(* IEC 61131-3 sources: 2026_Projet_YGO_ExcavatriceDragage/CODE/MAIN, 13 files *)

(* ---- GVL_Global.st ---- *)
(* ═══════════════════════════════════════════════════════════════
   🌐 GVL_Global — Variables globales d'utilité générale
   ───────────────────────────────────────────────────────────────
   🎯 Rôle : Regrouper les signaux et horloges système partagés qui
      ne sont pas spécifiques à la logique de simulation ni raccordés
      à des calibrations persistantes.
   ═══════════════════════════════════════════════════════════════ *)
{attribute 'qualified_only'}
VAR_GLOBAL
    BlinkClock1Hz              : BOOL;          // Horloge 1Hz pour clignotements (IHM ou diagnostic)
END_VAR

(* ---- PRG_00_Inputs.st ---- *)
(* ═══════════════════════════════════════════════════════════════
   📥 PRG_00_Inputs — Acquisition et conditionnement des ENTRÉES (PROGRAMME)
   ───────────────────────────────────────────────────────────────
   📄 Doc : DOC/AF_Partie6_IO_Conditioning_v1.2.md §5
   ⚙️ Exécuté par la tâche PLC (Task Manager) en position 0.
   ✅ Expose ses sorties en VAR_OUTPUT (lecture seule pour le reste du code).
   ═══════════════════════════════════════════════════════════════ *)

PROGRAM PRG_00_Inputs
VAR_OUTPUT
    // ── 🛑 SÉCURITÉS COMMUNES (NC — repos=TRUE sain, FALSE=défaut/fil coupé) ──────────────
    // 🔧 REX 2026-07-07 : précision terrain — EmergencyStopOk_DI (retour contact auxiliaire NO)
    // est en fait la confirmation que le CONTACTEUR DE PUISSANCE est réellement engagé (1=actif),
    // PAS la boucle AU elle-même (ça, c'est EmergencyChainOK_DI, ci-dessous). Nom EmergencyStopOk
    // conservé tel quel (contrat FB standard Partie3 §1, utilisé partout) — reste le portail
    // maître du programme, car "puissance réellement présente" est la garantie la plus forte.
    EmergencyStopOk      : BOOL;   // 🚨 Contacteur de puissance confirmé engagé : TRUE=armé/actif ✅ | FALSE=non armé ou coupure 🔴
    EmergencyChain       : BOOL;   // 🔗 REX 2026-07-07 : boucle AU (coup-de-poing + contact PLC) : TRUE=saine ✅ | FALSE=AU appuyé ou PowerCutOff PLC actif 🔴 — précondition à l'armement, PAS le portail maître
    TopPositionSensor    : BOOL;   // 🔝 Fin de course HAUT (NC) : TRUE=libre ✅ | FALSE=butée atteinte 🔴→ForbidAscent
    SlackCableSwitch     : BOOL;   // 🔗 Mou câble sur tambour M2 (NC) : TRUE=câble tendu ✅ | FALSE=mou détecté 🔴→ForbidDescent
    PhaseRotationOk      : BOOL;   // ⚡ Rotation phases élec. (NC) : TRUE=phases OK ✅ | FALSE=inversées/absentes 🔴→SafeStop
    // 🆕 REX 2026-07-08 : retour thermique COMMUN aux 3 freins M1/M2/M3 (1 seul fil, impossible
    // de savoir lequel des 3 est en cause) — demande utilisateur : la perte de ce retour peut
    // signifier un frein qui colle instantanément (frein à manque de courant) → traité comme
    // les autres défauts francs du domaine, escalade PowerCutOff côté FB_Safety_Winch/_Chariot
    // (voir bit10/bit3 respectifs).
    BrakeThermalFeedback : BOOL;   // 🌡️ Thermique frein M1/M2/M3 commun (NC) : TRUE=temp OK ✅ | FALSE=surchauffe ou coupure 🔴→SafeStop+PowerCutOff

    // ── 🪝 TREUIL M1 (frein=NC ; feedback contacteurs=retour unique REX 2026-07-07) ─────
    M1FwdRevSpeedFeedbackOff : BOOL; // 📡 REX 2026-07-07 : retour unique "tous contacteurs (sens+vitesse)
                                      // retombés" M1 — remplace M1ContactorFeedbackFwd/Rev (feedback
                                      // individuel par sens supprimé côté matériel, plus jamais câblé).
                                      // TRUE = tous retombés (sain, rien d'engagé)
    M1ThermalFeedback      : BOOL; // 🌡️ Thermique moteur M1 (NC) : TRUE=temp OK ✅ | FALSE=surchauffe ou coupure 🔴
    M1BrakeFeedback        : BOOL; // 🔒 Retour frein M1 (NC) : TRUE=frein serré repos ✅ | FALSE=desserré/coupure 🔴

    // ── 🪝 TREUIL M2 (même logique que M1) ──────────────────────────────────────────────
    M2FwdRevSpeedFeedbackOff : BOOL; // 📡 REX 2026-07-07 : idem M1, voir ci-dessus
    M2ThermalFeedback      : BOOL; // 🌡️ Thermique moteur M2 (NC) : TRUE=surchauffe ou coupure 🔴→SafeStop+PowerCutOff
    M2BrakeFeedback        : BOOL; // 🔒 Retour frein M2 (NC) : TRUE=serré repos ✅ | FALSE=desserré/coupure 🔴

    // ── ↔️ CHARIOT M3 (capteurs position=NO — position atteinte=TRUE) ────────────────────
    ChariotPosFosse1      : BOOL;  // 📍 Position fosse 1 (NO) : TRUE=chariot en fosse 1 ✅ | FALSE=absent
    ChariotPosFosse2      : BOOL;  // 📍 Position fosse 2 (NO) : TRUE=chariot en fosse 2 ✅ | FALSE=absent
    ChariotPosMaintenance : BOOL;  // 🔧 Position maintenance (NO) : TRUE=en position service ✅ | FALSE=absent
    ChariotPosTremie      : BOOL;  // 🗑️ Position trémie vidange (NO) : TRUE=en position trémie ✅ | FALSE=absent
    M3BrakeFeedback       : BOOL;  // 🔒 Retour frein chariot M3 (NC) : TRUE=serré repos ✅ | FALSE=desserré 🔴

    // 🆕 Variables intermédiaires filtrées/simulées pour contourner la lecture seule des PDO
    M3_StatusWord_Filtered        : WORD;
    M3_ActualFrequencyHz_Filtered : UINT;
END_VAR
VAR
    // Instances de filtrage
    instEmergencyStopOk   : FB_Input;
    instEmergencyChain    : FB_Input; // 🔧 REX 2026-07-07
    instSlackCableSwitch  : FB_Input;
    instTopPositionSensor : FB_Input;
    instCtrlPhaseRotation : FB_Input;
    instBrakeThermalFeedback : FB_Input; // 🆕 REX 2026-07-08

    instM1FwdRevSpeedFeedbackOff : FB_Input; // 🔧 REX 2026-07-07 : remplace instM1ContactorFwd/Rev
    instM1Thermal      : FB_Input;
    instM1BrakeFeedback: FB_Input;

    instM2FwdRevSpeedFeedbackOff : FB_Input; // 🔧 REX 2026-07-07 : remplace instM2ContactorFwd/Rev
    instM2Thermal      : FB_Input;
    instM2BrakeFeedback: FB_Input;

    instChariotPosFosse1      : FB_Input;
    instChariotPosFosse2      : FB_Input;
    instChariotPosMaintenance : FB_Input;
    instChariotPosTremie      : FB_Input;
    instM3BrakeFeedback       : FB_Input;

    // 🧪 Simulation dynamique du trajet chariot M3 (Lot 4, non prioritaire — voir AF_Partie13)
    instSimChariot            : FB_Sim_Chariot;

    // 🧪 Simulation de la chaîne de sécurité AU / réarmement (Lot 1, combler le trou d'intégration)
    instSimSafety             : FB_Sim_Safety;

    // 🧪 Simulation des retours contacteurs et freins M1/M2 (Lot 1)
    M1_FwdRevSpeedFeedbackOff_Simulated : BOOL;
    M1BrakeFeedback_Simulated           : BOOL;
    M2_FwdRevSpeedFeedbackOff_Simulated : BOOL;
    M2BrakeFeedback_Simulated           : BOOL;
    M3BrakeFeedback_Simulated           : BOOL;

    // 🆕 REX 2026-07-08 (4) : cohérence simulation capteur haut (voir instTopPositionSensor ci-dessous)
    SimTopSensorTriggered                : BOOL;
END_VAR

// === IMPLEMENTATION (corps du PROGRAM PRG_00_Inputs) ===

// 🛑 ─── COMMUN ────────────────────────────────────────────────────────────
// 🧪 Simulation : chaque OR ci-dessous force le capteur à son état "sain" (famille
// sécurité, TRUE=OK) quand SimulationModeActive ET que ce capteur précis n'est
// pas encore câblé réellement (GVL_Simulation.*_IsReal). Voir AF_Partie13.

// Simulation de la chaîne de sécurité AU / réarmement (Lot 1)
instSimSafety(
    Enable          := GVL_Simulation.SimulationModeActive AND NOT GVL_Simulation.EmergencyStopChain_IsReal,
    PowerCutOff_A   := PowerCutOff_A_RQ,
    PowerCutOff_B   := PowerCutOff_B_RQ,
    EmergencyArming := EmergencyArming_RQ
);

instEmergencyStopOk(InputRaw := EmergencyStopOk_DI OR instSimSafety.SimContactorOk, FilterTime := T#20MS);
EmergencyStopOk := instEmergencyStopOk.State;

// 🔧 REX 2026-07-07 : boucle AU (coup-de-poing + contact PLC) — distincte du contacteur de
// puissance ci-dessus. Réutilise le même flag simulation (même sous-système physique AU).
instEmergencyChain(InputRaw := EmergencyChainOK_DI OR instSimSafety.SimChainOk, FilterTime := T#20MS);
EmergencyChain := instEmergencyChain.State;

// 🔧 REX 2026-07-07 : M1_M2_SlackCableSwitch_DI → M2_SlackCableSwitch_DI (capteur physiquement
// uniquement sur le tambour M2, le préfixe M1_M2_ ne reflétait pas la réalité du câblage)
instSlackCableSwitch(InputRaw := M2_SlackCableSwitch_DI OR (GVL_Simulation.SimulationModeActive AND NOT GVL_Simulation.SlackCableSwitch_IsReal), FilterTime := T#20MS);
SlackCableSwitch := instSlackCableSwitch.State;

// 🆕 REX 2026-07-08 (4) : cohérence simulation (demande utilisateur) — l'ancien câblage forçait
// TopPositionSensor à TOUJOURS TRUE (sain) en simulation, quelle que soit la position codeur :
// impossible de tester bit5/Méca D (capteur haut) en simulation, il ne se déclenchait JAMAIS.
// Dérivé désormais de la position M1 simulée (référence de l'ensemble, voir FB_Grappin/
// ActiveOffsetM) — 1 cycle de retard (PRG_00 avant PRG_02 dans l'ordre de tâche), négligeable,
// même principe déjà assumé ailleurs (EncoderFaultPresent, GrappinHoldStillActive).
SimTopSensorTriggered := (NOT PRG_04_Modes.instModes.InhibitM1 AND (PRG_02_Encoders.instEncoderScaleM1.CablePosM >= GVL_PERSISTENT.HomingTargetM1_M))
                      OR (NOT PRG_04_Modes.instModes.InhibitM2 AND (PRG_02_Encoders.instEncoderScaleM2.CablePosM >= GVL_PERSISTENT.HomingTargetM2_M));
instTopPositionSensor(InputRaw := M1_M2_TopPositionSensor_DI OR (GVL_Simulation.SimulationModeActive AND NOT GVL_Simulation.TopPositionSensor_IsReal AND NOT SimTopSensorTriggered), FilterTime := T#20MS);
TopPositionSensor := instTopPositionSensor.State;

instCtrlPhaseRotation(InputRaw := CtrlPhaseRotation_DI OR (GVL_Simulation.SimulationModeActive AND NOT GVL_Simulation.PhaseRotationOk_IsReal), FilterTime := T#20MS);
PhaseRotationOk := instCtrlPhaseRotation.State;

// 🆕 REX 2026-07-08 : thermique frein commun M1/M2/M3 (1 seul fil, voir bandeau ci-dessus)
instBrakeThermalFeedback(InputRaw := BrakeThermalFeedback_DI OR (GVL_Simulation.SimulationModeActive AND NOT GVL_Simulation.BrakeThermal_IsReal), FilterTime := T#20MS);
BrakeThermalFeedback := instBrakeThermalFeedback.State;

// 🪝 ─── WINCH M1 ──────────────────────────────────────────────────────────
// 🧪 Simulation des retours contacteurs M1 (retombés si aucun sens/vitesse commandé)
M1_FwdRevSpeedFeedbackOff_Simulated := NOT (PRG_10_Outputs.M1RelayFwd OR PRG_10_Outputs.M1RelayRev OR PRG_10_Outputs.M1SpeedContactor1 OR PRG_10_Outputs.M1SpeedContactor2 OR PRG_10_Outputs.M1SpeedContactor3 OR PRG_10_Outputs.M1SpeedContactor4);
instM1FwdRevSpeedFeedbackOff(InputRaw := SEL(GVL_Simulation.SimulationModeActive AND NOT GVL_Simulation.ContactorFeedbackM1_IsReal, M1_FwdRevSpeedFeedbackOff_DI, M1_FwdRevSpeedFeedbackOff_Simulated), FilterTime := T#20MS);
M1FwdRevSpeedFeedbackOff := instM1FwdRevSpeedFeedbackOff.State;

instM1Thermal(InputRaw := M1_ThermalFeedback_DI OR (GVL_Simulation.SimulationModeActive AND NOT GVL_Simulation.ThermalM1_IsReal), FilterTime := T#20MS);
M1ThermalFeedback := instM1Thermal.State;

// 🧪 Simulation du retour frein M1 (fermé si commande inactive)
M1BrakeFeedback_Simulated := NOT PRG_10_Outputs.M1BrakeCmd;
instM1BrakeFeedback(InputRaw := SEL(GVL_Simulation.SimulationModeActive AND NOT GVL_Simulation.ContactorFeedbackM1_IsReal, M1_BrakeFeedback_DI, M1BrakeFeedback_Simulated), FilterTime := T#20MS);
M1BrakeFeedback := instM1BrakeFeedback.State;

// 🪝 ─── WINCH M2 ──────────────────────────────────────────────────────────
// 🧪 Simulation des retours contacteurs M2 (retombés si aucun sens/vitesse commandé)
M2_FwdRevSpeedFeedbackOff_Simulated := NOT (PRG_10_Outputs.M2RelayFwd OR PRG_10_Outputs.M2RelayRev OR PRG_10_Outputs.M2SpeedContactor1 OR PRG_10_Outputs.M2SpeedContactor2 OR PRG_10_Outputs.M2SpeedContactor3 OR PRG_10_Outputs.M2SpeedContactor4);
instM2FwdRevSpeedFeedbackOff(InputRaw := SEL(GVL_Simulation.SimulationModeActive AND NOT GVL_Simulation.ContactorFeedbackM2_IsReal, M2_FwdRevSpeedFeedbackOff_DI, M2_FwdRevSpeedFeedbackOff_Simulated), FilterTime := T#20MS);
M2FwdRevSpeedFeedbackOff := instM2FwdRevSpeedFeedbackOff.State;

instM2Thermal(InputRaw := M2_ThermalFeedback_DI OR (GVL_Simulation.SimulationModeActive AND NOT GVL_Simulation.ThermalM2_IsReal), FilterTime := T#20MS);
M2ThermalFeedback := instM2Thermal.State;

// 🧪 Simulation du retour frein M2 (fermé si commande inactive)
M2BrakeFeedback_Simulated := NOT PRG_10_Outputs.M2BrakeCmd;
instM2BrakeFeedback(InputRaw := SEL(GVL_Simulation.SimulationModeActive AND NOT GVL_Simulation.ContactorFeedbackM2_IsReal, M2_BrakeFeedback_DI, M2BrakeFeedback_Simulated), FilterTime := T#20MS);
M2BrakeFeedback := instM2BrakeFeedback.State;

// ↔️ ─── CHARIOT M3 ────────────────────────────────────────────────────────
// 🧪 Simulation dynamique du trajet M3 (FB_Sim_Chariot, non prioritaire — voir AF_Partie13
// §Chariot). Appelée AVANT les FB_Input pour que ses sorties soient à jour au même cycle
// (sinon décalage d'1 cycle sur le OR ci-dessous). Remplace le forçage manuel en vue instance.
// 🔧 REX 2026-07-15 (3) : RelayFwd/RelayRev câblés sur M3_CommandWord (variable globale
// mappée PDO EtherCAT, valeur réellement envoyée, Auto ET Manu confondus) — ex-
// GVL_Chariot_M3_Stub.M3_RelayFwd/Rev n'étaient plus jamais écrits depuis l'abandon du mode
// relais DEGRADED_IO (v0.4.11), la simulation de trajet M3 restait bloquée en permanence
// (relais toujours FALSE). Lecture décalée d'1 cycle (10ms, M3_CommandWord réécrit en position
// 10 par PRG_10_Outputs après ce PRG_00) — négligeable devant TravelTimeS (8s).
instSimChariot(
    Enable      := GVL_Simulation.SimulationModeActive AND NOT GVL_Simulation.ChariotPosition_IsReal,
    TargetNum   := GVL_Chariot_M3_Stub.StubChariotPositionSelect_IHM,
    RelayFwd    := M3_CommandWord = 1,
    RelayRev    := M3_CommandWord = 2,
    TravelTimeS := 8.0
);

instChariotPosFosse1(InputRaw := PosFosse1_DI OR instSimChariot.PosFosse1, FilterTime := T#20MS);
ChariotPosFosse1 := instChariotPosFosse1.State;

instChariotPosFosse2(InputRaw := PosFosse2_DI OR instSimChariot.PosFosse2, FilterTime := T#20MS);
ChariotPosFosse2 := instChariotPosFosse2.State;

instChariotPosMaintenance(InputRaw := PosMaintenance_DI OR instSimChariot.PosMaintenance, FilterTime := T#20MS);
ChariotPosMaintenance := instChariotPosMaintenance.State;

instChariotPosTremie(InputRaw := PosTremie_DI OR instSimChariot.PosTremie, FilterTime := T#20MS);
ChariotPosTremie := instChariotPosTremie.State;

// 🧪 Simulation du retour frein M3 (fermé/NC=TRUE si commande inactive)
M3BrakeFeedback_Simulated := NOT PRG_07_ChariotControl.instChariotM3.BrakeCmd;
instM3BrakeFeedback(InputRaw := SEL(GVL_Simulation.SimulationModeActive AND NOT GVL_Simulation.ContactorFeedbackM3_IsReal, M3_BrakeFeedback_DI, M3BrakeFeedback_Simulated), FilterTime := T#20MS);
M3BrakeFeedback := instM3BrakeFeedback.State;

// 🧪 Simulation/Filtrage des retours variateur EtherCAT M3 (lecture seule physique contournée)
IF GVL_Simulation.SimulationModeActive AND NOT GVL_Simulation.VariateurM3_IsReal THEN
    M3_ActualFrequencyHz_Filtered := M3_SetpointFrequencyHz;

    // Status Word : Bit0 (Operation), Bit7 (Operation Enable)
    IF M3_CommandWord = 1 THEN
        M3_StatusWord_Filtered := 16#0081; // Operation + Operation Enable
    ELSIF M3_CommandWord = 2 THEN
        M3_StatusWord_Filtered := 16#0089; // Operation + Operation Enable + Reverse (bit3)
    ELSE
        M3_StatusWord_Filtered := 16#0080; // Stopped + Operation Enable
    END_IF;
ELSE
    M3_ActualFrequencyHz_Filtered := M3_ActualFrequencyHz;
    M3_StatusWord_Filtered        := M3_StatusWord;
END_IF;

(* ---- PRG_01_Diagnostics.st ---- *)
(* ═══════════════════════════════════════════════════════════════
   📡 PRG_01_Diagnostics — États bus de terrain et Joystick (PROGRAMME)
   ───────────────────────────────────────────────────────────────
   ⚙️ Exécuté par la tâche PLC en position 1.
   ═══════════════════════════════════════════════════════════════ *)

PROGRAM PRG_01_Diagnostics
VAR
    instDiagCanOpen  : FB_DiagCanOpen;       // Diagnostic CAN/Joystick
    instDiagEthercat : FB_DiagEthercat;      // Diagnostic EtherCAT (3 devices)
    FB_Joystick_0    : FB_Joystick;          // Traitement joystick (calib/filtre/rampe)
    instSimJoystick  : FB_Sim_Joystick;      // 🧪 Simulation joystick (Lot 3 — voir CODE/SIMULATION/)
END_VAR

// === IMPLEMENTATION (corps du PROGRAM PRG_01_Diagnostics) ===

// 🧪 0. Simulation Joystick (Lot 3, priorité — voir CODE/SIMULATION/FB_Sim_Joystick.st) : appelée
// AVANT FB_Joystick_0 pour que ses sorties soient à jour au même cycle. Remplace l'ancien bypass
// homme-mort codé en dur dans FB_Joystick (GVL_DEBUG.DBG_DeadmanBypass_TEST) : quand
// NOT JoystickSignal_IsReal, ses sorties remplacent les entrées brutes ci-dessous ; le homme-mort
// réel de FB_Joystick n'est plus jamais contourné.
// 🆕 REX 2026-07-08 : gardé désormais par JoystickSignal_IsReal (PAS Joystick_IsReal, qui ne
// couvre que le bus CANopen ci-dessous) — granularité séparée demandée par l'utilisateur : tester
// le signal joystick réel sans dépendre du diagnostic bus/nœud CANopen (encore simulé sain).
instSimJoystick(
    Enable          := GVL_Simulation.SimulationModeActive AND NOT GVL_Simulation.JoystickSignal_IsReal,
    NeutralRaw      := GVL_Simulation.JoystickForceNeutralRaw,
    MaxRaw          := GVL_Simulation.JoystickForceMaxRaw
);

// 1. Diagnostics CANopen — 🆕 REX 2026-07-08 : gardé par Joystick_IsReal UNIQUEMENT (bus/nœud),
// indépendant de JoystickSignal_IsReal (signal brut ci-dessus) — granularité séparée.
instDiagCanOpen(
    Enable := TRUE,
    Reset := PRG_09_Supervision.FaultMachineReset_IHM,
    CanOnline := (CANbus.GetBusState() = 1) OR (GVL_Simulation.SimulationModeActive AND NOT GVL_Simulation.Joystick_IsReal), // 1 = ACTIVE (ou simulation)
    CanOperational := (JOY1_JOYSTICK_MCB560_CO4201A.GetDeviceState() = DEVICE_STATE.RUNNING) OR (GVL_Simulation.SimulationModeActive AND NOT GVL_Simulation.Joystick_IsReal)
);

// 2. Diagnostics EtherCAT (variateur + 2 codeurs)
instDiagEthercat(
    Enable := TRUE,
    Reset := PRG_09_Supervision.FaultMachineReset_IHM,          // 🔑 Bouton général machine
    VariateurWcState := (AC600_ECAT_Drive.GetDeviceState() <> DEVICE_STATE.RUNNING) AND NOT (GVL_Simulation.SimulationModeActive AND NOT GVL_Simulation.VariateurM3_IsReal),
    VariateurSlaveState := SEL((GVL_Simulation.SimulationModeActive AND NOT GVL_Simulation.VariateurM3_IsReal) OR (AC600_ECAT_Drive.GetDeviceState() = DEVICE_STATE.RUNNING), 0, 8),
    EncoderM1WcState := (COD1_CODEUR.GetDeviceState() <> DEVICE_STATE.RUNNING) AND NOT (GVL_Simulation.SimulationModeActive AND NOT GVL_Simulation.EncoderM1_IsReal),
    EncoderM1SlaveState := SEL((GVL_Simulation.SimulationModeActive AND NOT GVL_Simulation.EncoderM1_IsReal) OR (COD1_CODEUR.GetDeviceState() = DEVICE_STATE.RUNNING), 0, 8),
    EncoderM2WcState := (COD2_CODEUR.GetDeviceState() <> DEVICE_STATE.RUNNING) AND NOT (GVL_Simulation.SimulationModeActive AND NOT GVL_Simulation.EncoderM2_IsReal),
    EncoderM2SlaveState := SEL((GVL_Simulation.SimulationModeActive AND NOT GVL_Simulation.EncoderM2_IsReal) OR (COD2_CODEUR.GetDeviceState() = DEVICE_STATE.RUNNING), 0, 8)
);

// 3. Acquisition Joystick — RawX/RawY/RawButton simulés (instSimJoystick) quand NOT JoystickSignal_IsReal
// 🔴🔧 REX 2026-07-07 — TEST BANC UNIQUEMENT, PAS DE VALEUR PRODUCTION :
//    DeadmanRearmTimeout 10s → 5min, NeutralHoldTime 500ms → 1s (confort d'essai, moins de
//    réappuis/traversées à gérer). ⚠️ RÉDUIT RÉELLEMENT LA SÉCURITÉ HOMME-MORT — à repasser
//    impérativement à T#10S / T#500MS (ou retirer ces 2 lignes, le FB reprend ses défauts sûrs)
//    avant toute mise en service réelle avec la machine.
FB_Joystick_0(
    Enable              := TRUE,
    EmergencyStopOk     := PRG_00_Inputs.EmergencyStopOk,
    Reset               := PRG_09_Supervision.FaultMachineReset_IHM,
    Mode                := PRG_04_Modes.instModes.Mode,  // 🆕 REX 2026-07-08 : désarme le homme-mort au changement de mode
    // 🆕 REX 2026-07-08 : PRG_01 (position 1) s'exécute AVANT PRG_06 (position 6) — GrappinBusy lu
    // ici reflète donc le Busy du scan PRÉCÉDENT (retard d'1 scan, ~10ms, sur la détection du front
    // descendant). Sans impact pratique : très inférieur aux temps de réponse frein/contacteurs
    // (100-300ms, voir FB_Brake) — la commande n'a pas le temps de produire un mouvement réel.
    GrappinBusy         := PRG_06_WinchControl.instGrappin.Busy,
    NeutralXMem         := GVL_PERSISTENT.JoystickNeutralX,
    NeutralYMem         := GVL_PERSISTENT.JoystickNeutralY,
    BusCanOpenOP        := instDiagCanOpen.busCanOpen,
    JoystickOP          := instDiagCanOpen.Joystick,
    RawX                := SEL(instSimJoystick.Enable, JoyXRaw_ANA1, instSimJoystick.RawX),
    RawY                := SEL(instSimJoystick.Enable, JoyYRaw_ANA2, instSimJoystick.RawY),
    RawButton           := SEL(instSimJoystick.Enable, JoyBtnRaw, instSimJoystick.RawButton),
    Calibrate           := GVL_IHM.JoystickJOY1.Calibrate,
    InvertX             := FALSE,
    InvertY             := FALSE,
    Deadband            := 10.0,
    FilterTime          := TIME#100ms,
    AccelRate           := 50.0,
    DecelRate           := 150.0,
    // 🛡️ Délais de sécurité Homme-Mort : temporisations courtes (10s/500ms) si joystick réel, longues (5min/1s) si simulé
    DeadmanRearmTimeout := SEL(NOT GVL_Simulation.SimulationModeActive OR GVL_Simulation.JoystickSignal_IsReal, T#5M, T#10S),
    NeutralHoldTime     := SEL(NOT GVL_Simulation.SimulationModeActive OR GVL_Simulation.JoystickSignal_IsReal, T#1S, T#500MS)
);

(* ---- PRG_02_Encoders.st ---- *)
(* ═══════════════════════════════════════════════════════════════
   🧲 PRG_02_Encoders — Acquisition, Recalage (Homing) et Sécurité Codeurs
   ───────────────────────────────────────────────────────────────
   ⚙️ Exécuté par la tâche PLC en position 2.
   ✅ Expose ses défauts en VAR_OUTPUT (1 cycle de retard assumé pour instModes).
   ═══════════════════════════════════════════════════════════════ *)

PROGRAM PRG_02_Encoders
VAR_OUTPUT
    EncoderFaultPresent   : BOOL;   // OR des deux - lu par PRG_04_Modes au cycle suivant
    EncoderFaultPresentM1 : BOOL;
    EncoderFaultPresentM2 : BOOL;
END_VAR
VAR
    // 🧪 Simulation banc de test (Lot 2 — voir CODE/SIMULATION/FB_Sim_Encoder.st)
    instSimEncoderM1      : FB_Sim_Encoder;
    instSimEncoderM2      : FB_Sim_Encoder;
    M1_RawPosToUse        : UDINT;
    M2_RawPosToUse        : UDINT;

    // Instances
    instEncoderAbsM1   : FB_Encoder_Abs;
    instEncoderScaleM1 : FB_Encoder_Scale;
    instHomingM1       : FB_Encoder_Homing;
    instEncoderAbsM2   : FB_Encoder_Abs;
    instEncoderScaleM2 : FB_Encoder_Scale;
    instHomingM2       : FB_Encoder_Homing;
    instEncoderSafetyM1 : FB_Encoder_Safety;
    instEncoderSafetyM2 : FB_Encoder_Safety;

    M1_SimSpeedPct      : REAL;
    M2_SimSpeedPct      : REAL;
    M1_IsReal           : BOOL;         // ⚡ Indique si le treuil M1 est configuré comme réel
    M2_IsReal           : BOOL;         // ⚡ Indique si le treuil M2 est configuré comme réel
END_VAR

// === IMPLEMENTATION (corps du PROGRAM PRG_02_Encoders) ===

// 🆕 Détermination de la réalité des treuils (Conditional Bypass Doctrine)
M1_IsReal := NOT GVL_Simulation.SimulationModeActive OR GVL_Simulation.EncoderM1_IsReal OR GVL_Simulation.ContactorFeedbackM1_IsReal OR GVL_Simulation.ThermalM1_IsReal;
M2_IsReal := NOT GVL_Simulation.SimulationModeActive OR GVL_Simulation.EncoderM2_IsReal OR GVL_Simulation.ContactorFeedbackM2_IsReal OR GVL_Simulation.ThermalM2_IsReal;

// 🔧 REX 2026-07-15 (4) — CORRECTIF COMPILATION : ex-SEL(ManuActive, ...) référençait
// PRG_10_Outputs.SpeedRefPct, supprimé lors du passage de Manu sur FB_Winch (REX 2026-07-15 (2)).
// Plus besoin de distinguer Auto/Manu ici : instWinchM1/M2.SpeedRamp.Current est désormais LA
// vitesse rampée réelle dans les DEUX cas (FB_Winch pilote M1/M2 qu'on soit en Auto ou en Manu).
M1_SimSpeedPct := PRG_06_WinchControl.instWinchM1.SpeedRamp.Current;
M2_SimSpeedPct := PRG_06_WinchControl.instWinchM2.SpeedRamp.Current;

// 1. SIMULATION SUR BANC DE TEST (Lot 2, granularité indépendante M1/M2 — voir AF_Partie13)
// 🔧 REX 2026-07-08 : RawPos (VAR_IN_OUT) référence GVL_PERSISTENT.SimEncoderRawPosM1/M2 —
// survit à un reset froid comme le ferait un vrai codeur absolu physique (voir GVL_PERSISTENT.st).
instSimEncoderM1(
    Enable      := GVL_Simulation.SimulationModeActive AND NOT GVL_Simulation.EncoderM1_IsReal,
    // 🔧 REX 2026-07-15 (2) : lit directement instWinchM1 (PRG_06_WinchControl) — M1 est désormais
    // piloté par FB_Winch en Auto ET en Manu (ex-SimM1Fwd_Eff/PRG_10_Outputs retiré, obsolète) :
    // RelayFwd/RelayRev respectent déjà SafeStop/ForbidAscent/ForbidDescent nativement, plus besoin
    // de signaux Sim dédiés.
    RelayFwd    := PRG_06_WinchControl.instWinchM1.RelayFwd,
    RelayRev    := PRG_06_WinchControl.instWinchM1.RelayRev,
    SpeedRefPct := M1_SimSpeedPct,
    PresetCmd   := (COD1_PresettTrigCmd = 2),
    PresetValue := COD1_PresetValue,
    SpeedScaleFactor := GVL_Simulation.EncoderSimSpeedFactor,  // 🔧 REX 2026-07-07 : confort de test
    // 🆕 REX 2026-07-08 (4) : injection saut de test (Concept 1 / Méca E) — 4096 = PointsPerRev/CableM_PerRev (8192/2.0)
    TestOffsetCmd := GVL_Simulation.InjectSyncDeviationM1,
    TestOffsetPts := REAL_TO_DINT(GVL_Simulation.SyncDeviationOffsetM * 4096.0),
    RawPos      := GVL_PERSISTENT.SimEncoderRawPosM1
);
instSimEncoderM2(
    Enable      := GVL_Simulation.SimulationModeActive AND NOT GVL_Simulation.EncoderM2_IsReal,
    // 🔧 REX 2026-07-15 (2) : idem M1 ci-dessus, lit instWinchM2 (ex-SimM2Fwd_Eff retiré).
    RelayFwd    := PRG_06_WinchControl.instWinchM2.RelayFwd,
    RelayRev    := PRG_06_WinchControl.instWinchM2.RelayRev,
    SpeedRefPct := M2_SimSpeedPct,
    PresetCmd   := (COD2_PresettTrigCmd = 2),
    PresetValue := COD2_PresetValue,
    SpeedScaleFactor := GVL_Simulation.EncoderSimSpeedFactor,  // 🔧 REX 2026-07-07 : confort de test
    // 🆕 REX 2026-07-08 (4) : injection saut de test (Concept 1 / Méca E)
    TestOffsetCmd := GVL_Simulation.InjectSyncDeviationM2,
    TestOffsetPts := REAL_TO_DINT(GVL_Simulation.SyncDeviationOffsetM * 4096.0),
    RawPos      := GVL_PERSISTENT.SimEncoderRawPosM2
);

// Aiguillage (par device — 🔧 REX 2026-07-07 : ne PAS utiliser Operational, forcé à TRUE en
// simulation par PRG_01_Diagnostics [SEL sur EncoderMx_IsReal] pour ne pas remonter de faux
// défaut bus — ça sélectionnait donc systématiquement COD1/COD2_PosValue [réel, figé à 0] au
// lieu de la position simulée, bloquant tout homing/mouvement testé en simulation.
IF (GVL_Simulation.SimulationModeActive AND NOT GVL_Simulation.EncoderM1_IsReal) THEN
    M1_RawPosToUse := instSimEncoderM1.RawPosOut;
ELSE
    M1_RawPosToUse := COD1_PosValue;
END_IF;

IF (GVL_Simulation.SimulationModeActive AND NOT GVL_Simulation.EncoderM2_IsReal) THEN
    M2_RawPosToUse := instSimEncoderM2.RawPosOut;
ELSE
    M2_RawPosToUse := COD2_PosValue;
END_IF;

// 2. TREUIL M1 (Abs → Homing → Scale)
// 🔧 REX 2026-07-07 : Homing appelé AVANT Scale (et non l'inverse) — Scale lit HomingRefRaw en
// entrée ; si Scale s'exécutait avant Homing, un homing réussi au cycle N ne serait répercuté
// sur CablePosM qu'au cycle N+1, alors que instHomingM1.Busy (→ InReferencingMode côté
// FB_Safety_Winch) retombe dès le cycle N — décalage d'1 cycle qui désynchronise le garde-fou
// anti-transition de Méca A (bit7) et provoque un faux déclenchement PowerCutOff au cycle N+1
// (saut de position vu hors fenêtre "référencement en cours"). Homing ne dépend d'aucune sortie
// de Scale (RawPos vient d'instEncoderAbsM1) : aucune dépendance circulaire, réordonnancement sûr.
instEncoderAbsM1(
    Enable              := TRUE,
    Reset               := PRG_09_Supervision.FaultMachineReset_IHM,
    EmergencyStopOk     := PRG_00_Inputs.EmergencyStopOk,
    Mode                := PRG_04_Modes.instModes.Mode,
    RawPosIn            := M1_RawPosToUse,
    AlarmsIn            := SEL(instSimEncoderM1.Enable, COD1_Alarms, 0),
    WarningsIn          := SEL(instSimEncoderM1.Enable, COD1_Warnings, 0),
    SlaveOperational    := PRG_01_Diagnostics.instDiagEthercat.EncoderM1.Operational OR instSimEncoderM1.Enable,
    PresetRequest       := instHomingM1.PresetRequest OR (PRG_10_Outputs.ManuActive AND NOT M1_IsReal AND GVL_IHM.IHM_MANU.HomingEncoder_M1),
    PresetValue         := SEL(PRG_10_Outputs.ManuActive AND NOT M1_IsReal AND GVL_IHM.IHM_MANU.HomingEncoder_M1, instHomingM1.PresetValue, 16777216)
);
COD1_PresettTrigCmd := instEncoderAbsM1.PresetTriggerCmd;
COD1_CodeSeqTrigCmd := instEncoderAbsM1.CodeSeqTriggerCmd;
COD1_PresetValue    := instEncoderAbsM1.PresetValueOut;

instHomingM1(
    Enable               := TRUE,
    Calib                := GVL_PERSISTENT.CalibM1,
    Reset                := PRG_09_Supervision.FaultMachineReset_IHM,
    EmergencyStopOk      := PRG_00_Inputs.EmergencyStopOk,
    Mode                 := PRG_04_Modes.instModes.Mode,
    // ─────────  Début modification IHM_MANU  ─────────
    // 🆕 REX 2026-07-09 : OR avec HomingEncoder_M1 (mise en service urgence) — même FB, mêmes
    // conditions de sécurité (Mode MAINT_N1/N2, arrêt confirmé), aucune nouvelle dérogation.
    Home                 := GVL_IHM.WinchM1.CmdHome OR GVL_IHM.IHM_MANU.HomingEncoder_M1, // 🔧 REX 2026-07-07 : fusion GVL_Encoder_Stub → GVL_IHM
    // ─────────  Fin modification IHM_MANU  ─────────
    ConfirmCoherence     := GVL_IHM.WinchM1.ConfirmCoherence, // 🔧 REX 2026-07-07 : fusion GVL_Encoder_Stub → GVL_IHM
    TopPositionSensor    := PRG_00_Inputs.TopPositionSensor,
    TopSensorPositionM   := GVL_PERSISTENT.HomingTargetM1_M,
    FwdRevSpeedFeedbackOff := PRG_00_Inputs.M1FwdRevSpeedFeedbackOff, // 🔧 REX 2026-07-07
    BrakeFeedback        := PRG_00_Inputs.M1BrakeFeedback,
    RawPos               := instEncoderAbsM1.RawPos,
    EncoderAvailable     := instEncoderAbsM1.EncoderAvailable,
    PresetAck            := instEncoderAbsM1.PresetAck,
    PresetNak            := instEncoderAbsM1.PresetNak,
    PointsPerRev         := 8192,
    MultiTurnRevsMax     := 4096,
    CableM_PerRev        := 2.0
);

instEncoderScaleM1(
    RawPos          := instEncoderAbsM1.RawPos,
    HomingRefRaw    := instHomingM1.HomingRefRaw,
    CableM_PerRev   := 2.0,
    PointsPerRev    := 8192
);

// 3. TREUIL M2 (Abs → Homing → Scale)
instEncoderAbsM2(
    Enable              := TRUE,
    Reset               := PRG_09_Supervision.FaultMachineReset_IHM,
    EmergencyStopOk     := PRG_00_Inputs.EmergencyStopOk,
    Mode                := PRG_04_Modes.instModes.Mode,
    RawPosIn            := M2_RawPosToUse,
    AlarmsIn            := SEL(instSimEncoderM2.Enable, COD2_Alarms, 0),
    WarningsIn          := SEL(instSimEncoderM2.Enable, COD2_Warnings, 0),
    SlaveOperational    := PRG_01_Diagnostics.instDiagEthercat.EncoderM2.Operational OR instSimEncoderM2.Enable,
    PresetRequest       := instHomingM2.PresetRequest OR (PRG_10_Outputs.ManuActive AND NOT M2_IsReal AND GVL_IHM.IHM_MANU.HomingEncoder_M2),
    PresetValue         := SEL(PRG_10_Outputs.ManuActive AND NOT M2_IsReal AND GVL_IHM.IHM_MANU.HomingEncoder_M2, instHomingM2.PresetValue, 16777216)
);
COD2_PresettTrigCmd := instEncoderAbsM2.PresetTriggerCmd;
COD2_CodeSeqTrigCmd := instEncoderAbsM2.CodeSeqTriggerCmd;
COD2_PresetValue    := instEncoderAbsM2.PresetValueOut;

instHomingM2(
    Enable               := TRUE,
    Calib                := GVL_PERSISTENT.CalibM2,
    Reset                := PRG_09_Supervision.FaultMachineReset_IHM,
    EmergencyStopOk      := PRG_00_Inputs.EmergencyStopOk,
    Mode                 := PRG_04_Modes.instModes.Mode,
    // ─────────  Début modification IHM_MANU  ─────────
    // 🆕 REX 2026-07-09 : OR avec HomingEncoder_M2 (mise en service urgence) — même FB, mêmes
    // conditions de sécurité (Mode MAINT_N1/N2, arrêt confirmé), aucune nouvelle dérogation.
    Home                 := GVL_IHM.WinchM2.CmdHome OR GVL_IHM.IHM_MANU.HomingEncoder_M2, // 🔧 REX 2026-07-07 : fusion GVL_Encoder_Stub → GVL_IHM
    // ─────────  Fin modification IHM_MANU  ─────────
    ConfirmCoherence     := GVL_IHM.WinchM2.ConfirmCoherence, // 🔧 REX 2026-07-07 : fusion GVL_Encoder_Stub → GVL_IHM
    TopPositionSensor    := PRG_00_Inputs.TopPositionSensor,
    TopSensorPositionM   := GVL_PERSISTENT.HomingTargetM2_M,
    FwdRevSpeedFeedbackOff := PRG_00_Inputs.M2FwdRevSpeedFeedbackOff, // 🔧 REX 2026-07-07
    BrakeFeedback        := PRG_00_Inputs.M2BrakeFeedback,
    RawPos               := instEncoderAbsM2.RawPos,
    EncoderAvailable     := instEncoderAbsM2.EncoderAvailable,
    PresetAck            := instEncoderAbsM2.PresetAck,
    PresetNak            := instEncoderAbsM2.PresetNak,
    PointsPerRev         := 8192,
    MultiTurnRevsMax     := 4096,
    CableM_PerRev        := 2.0
);

instEncoderScaleM2(
    RawPos          := instEncoderAbsM2.RawPos,
    HomingRefRaw    := instHomingM2.HomingRefRaw,
    CableM_PerRev   := 2.0,
    PointsPerRev    := 8192
);

// 4. SÉCURITÉ DE BORNAGE ET INCOHÉRENCE
instEncoderSafetyM1(
    Enable          := TRUE,
    Reset           := PRG_09_Supervision.FaultMachineReset_IHM,
    EmergencyStopOk := PRG_00_Inputs.EmergencyStopOk,
    Mode            := PRG_04_Modes.instModes.Mode,
    CablePosM       := instEncoderScaleM1.CablePosM,
    HomingSuspect   := instHomingM1.HomingSuspect,
    PositionMinM    := -99.0,
    PositionMaxM    := 99.0
);
EncoderFaultPresentM1 := instEncoderSafetyM1.EncoderIncoherent;

instEncoderSafetyM2(
    Enable          := TRUE,
    Reset           := PRG_09_Supervision.FaultMachineReset_IHM,
    EmergencyStopOk := PRG_00_Inputs.EmergencyStopOk,
    Mode            := PRG_04_Modes.instModes.Mode,
    CablePosM       := instEncoderScaleM2.CablePosM,
    HomingSuspect   := instHomingM2.HomingSuspect,
    PositionMinM    := -99.0,
    PositionMaxM    := 99.0
);
EncoderFaultPresentM2 := instEncoderSafetyM2.EncoderIncoherent;

EncoderFaultPresent := EncoderFaultPresentM1 OR EncoderFaultPresentM2;

// ─────────  Début modification IHM_MANU  ─────────
// 🎯 Référencement direct (bypass sécurité et modes) si HomingEncoder_M1/M2 activés en Manu (uniquement si SIMULÉ)
// Sinon, si les treuils sont réels, on utilise le homing normal sécurisé, et on réinitialise le bouton HMI dès que homing ok/erreur.
IF PRG_10_Outputs.ManuActive THEN
    IF GVL_IHM.IHM_MANU.HomingEncoder_M1 THEN
        IF NOT M1_IsReal THEN
            IF instEncoderAbsM1.PresetAck THEN
                GVL_PERSISTENT.CalibM1.HomingRefRaw := 16726016; // 16777216 - (12.5 * 8192 / 2.0)
                GVL_PERSISTENT.CalibM1.Homed := TRUE;
                GVL_PERSISTENT.CalibM1.HomingSuspect := FALSE;
                GVL_PERSISTENT.CalibM1.LastKnownRawPos := 16777216;
                GVL_IHM.IHM_MANU.HomingEncoder_M1 := FALSE; // Reset bouton HMI
            ELSIF instEncoderAbsM1.PresetNak THEN
                GVL_IHM.IHM_MANU.HomingEncoder_M1 := FALSE;
            END_IF;
        ELSE
            IF instEncoderAbsM1.PresetAck OR instHomingM1.Homed THEN
                GVL_IHM.IHM_MANU.HomingEncoder_M1 := FALSE;
            ELSIF instEncoderAbsM1.PresetNak OR instHomingM1.Error THEN
                GVL_IHM.IHM_MANU.HomingEncoder_M1 := FALSE;
            END_IF;
        END_IF;
    END_IF;

    IF GVL_IHM.IHM_MANU.HomingEncoder_M2 THEN
        IF NOT M2_IsReal THEN
            IF instEncoderAbsM2.PresetAck THEN
                GVL_PERSISTENT.CalibM2.HomingRefRaw := 16726016; // 16777216 - (12.5 * 8192 / 2.0)
                GVL_PERSISTENT.CalibM2.Homed := TRUE;
                GVL_PERSISTENT.CalibM2.HomingSuspect := FALSE;
                GVL_PERSISTENT.CalibM2.LastKnownRawPos := 16777216;
                GVL_IHM.IHM_MANU.HomingEncoder_M2 := FALSE; // Reset bouton HMI
            ELSIF instEncoderAbsM2.PresetNak THEN
                GVL_IHM.IHM_MANU.HomingEncoder_M2 := FALSE;
            END_IF;
        ELSE
            IF instEncoderAbsM2.PresetAck OR instHomingM2.Homed THEN
                GVL_IHM.IHM_MANU.HomingEncoder_M2 := FALSE;
            ELSIF instEncoderAbsM2.PresetNak OR instHomingM2.Error THEN
                GVL_IHM.IHM_MANU.HomingEncoder_M2 := FALSE;
            END_IF;
        END_IF;
    END_IF;
END_IF;
// ─────────  Fin modification IHM_MANU  ─────────

(* ---- PRG_03_Safety.st ---- *)
(* ═══════════════════════════════════════════════════════════════
   🛡️ PRG_03_Safety — Centralisation des surveillances et blocs Safety
   ───────────────────────────────────────────────────────────────
   ⚙️ Exécuté par la tâche PLC en position 3.
   ═══════════════════════════════════════════════════════════════ *)

PROGRAM PRG_03_Safety
VAR
    instSafetyWinchM1   : FB_Safety_Winch;
    instSafetyWinchM2   : FB_Safety_Winch;
    instSafetyChariotM3 : FB_Safety_Chariot;
END_VAR

// === IMPLEMENTATION (corps du PROGRAM PRG_03_Safety) ===

// 1. Sécurité Treuil M1
instSafetyWinchM1(
    // 🔧 REX 2026-07-15 (2) — SIMPLIFICATION : IHM_MANU pilote désormais M1 via FB_Winch
    // (PRG_06_WinchControl), qui a BESOIN d'un SafeStop/ForbidAscent/ForbidDescent réels pour
    // rampé/ralentir proprement (ex-doctrine "Conditional Bypass" devenue obsolète et RETIRÉE
    // ici : chaque capteur/retour a DÉJÀ sa propre granularité réel/simulé — GVL_Simulation.
    // EncoderM1_IsReal, ContactorFeedbackM1_IsReal, ThermalM1_IsReal, TopPositionSensor_IsReal,
    // SlackCableSwitch_IsReal — un composant simulé est déjà forcé "sain" en amont (PRG_00_Inputs/
    // PRG_02_Encoders), donc Enable n'a plus besoin de bypasser tout le domaine : un vrai défaut
    // sur un composant RÉEL protège, un composant SIMULÉ ne fait jamais défaut de lui-même).
    Enable              := NOT PRG_04_Modes.instModes.InhibitM1, // 🆕 REX 2026-07-08 : Inhibit (MAINT_N2) uniquement
    Reset               := PRG_09_Supervision.FaultMachineReset_IHM,
    EmergencyStopOk     := PRG_00_Inputs.EmergencyStopOk,
    Mode                := PRG_04_Modes.instModes.Mode,
    SyncEnable          := PRG_04_Modes.instModes.SyncEnable,
    JoystickOnline      := PRG_01_Diagnostics.instDiagCanOpen.Joystick.Online,
    JoystickOperational := PRG_01_Diagnostics.instDiagCanOpen.Joystick.Operational,
    EncoderAvailable    := PRG_02_Encoders.instEncoderAbsM1.EncoderAvailable,
    ThermalFeedback     := NOT PRG_00_Inputs.M1ThermalFeedback,
    BrakeThermalFeedback := NOT PRG_00_Inputs.BrakeThermalFeedback, // 🆕 REX 2026-07-08 — commun M1/M2/M3
    SlackCableDetected  := NOT PRG_00_Inputs.SlackCableSwitch,
    PhaseRotationOk     := PRG_00_Inputs.PhaseRotationOk,
    TopPositionSensor   := PRG_00_Inputs.TopPositionSensor,
    InReferencingMode   := PRG_02_Encoders.instHomingM1.Busy,
    CablePosM           := PRG_02_Encoders.instEncoderScaleM1.CablePosM,
    CableLimitDescentM  := GVL_PERSISTENT.CableLimitDescentM1_M,
    Direction           := PRG_06_WinchControl.M1_Direction_Active,
    Homed               := PRG_02_Encoders.instHomingM1.Homed,
    HomingSuspect       := PRG_02_Encoders.instHomingM1.HomingSuspect,
    TopLimitM           := GVL_PERSISTENT.HomingTargetM1_M,
    // 🔧 REX 2026-07-07 — Méca A/B/C (voir FB_Safety_Winch bandeau en-tête)
    FwdRevSpeedFeedbackOff := PRG_00_Inputs.M1FwdRevSpeedFeedbackOff,
    BrakeFeedback          := PRG_00_Inputs.M1BrakeFeedback,
    // 🔧 REX 2026-07-15 (7) — BUG CORRIGÉ (retour terrain, SafetyErrorId=256/bit8) : Méca B ne
    // regardait QUE le joystick CANopen pour détecter "commande opérateur" — en IHM_MANU piloté
    // par BOUTONS HMI (JoystickSelect=FALSE), le joystick reste au neutre en permanence, donc
    // MecaB_NoOperatorCmd restait TRUE en continu même pendant un mouvement légitime aux boutons
    // → SafeStop après PostRampTimeout (3s) dès qu'un mouvement HMI dépassait ce délai. Ajout des
    // boutons IHM_MANU bruts (M1 individuel + Couplé) — reste indépendant de l'arbitrage
    // PRG_06/FB_Winch (défense en profondeur intacte, lecture directe des boutons IHM comme le
    // joystick l'était déjà).
    JoystickYNeutral       := (ABS(PRG_01_Diagnostics.FB_Joystick_0.AxisCmdY.SpeedRef) < 0.1)
                              AND NOT GVL_IHM.IHM_MANU.M1_RelayFwd AND NOT GVL_IHM.IHM_MANU.M1_RelayRev
                              AND NOT GVL_IHM.IHM_MANU.M1_M2_RelayFwd AND NOT GVL_IHM.IHM_MANU.M1_M2_RelayRev,
    GrappinHoldStillActive := PRG_06_WinchControl.instGrappin.Busy, // Méca C — M1 doit rester immobile pendant le
                                                                     // grappin ; 1 cycle de retard accepté (PRG_03
                                                                     // avant PRG_06 dans l'ordre de tâche), négligeable
    // 🆕 REX 2026-07-08 (4) — Méca E : M2 corrigé de l'offset grappin actif (0 si grappin absent/ouvert),
    // ramené dans le référentiel M1 — comparaison valable quel que soit l'état du grappin
    ExpectedOtherWinchPosM := PRG_02_Encoders.instEncoderScaleM2.CablePosM - PRG_06_WinchControl.instGrappin.ActiveOffsetM,
    GrappinBusy            := PRG_06_WinchControl.instGrappin.Busy,
    CriticalSyncToleranceM := GVL_PERSISTENT.WinchCriticalSyncTolerance_M,
    OtherWinchInhibited    := PRG_04_Modes.instModes.InhibitM2 // 🆕 REX 2026-07-08 (7)
);

// 2. Sécurité Treuil M2
instSafetyWinchM2(
    // 🔧 REX 2026-07-15 (2) — même simplification que M1 ci-dessus (voir bandeau instSafetyWinchM1).
    Enable              := NOT PRG_04_Modes.instModes.InhibitM2, // 🆕 REX 2026-07-08 : Inhibit (MAINT_N2) uniquement
    Reset               := PRG_09_Supervision.FaultMachineReset_IHM,
    EmergencyStopOk     := PRG_00_Inputs.EmergencyStopOk,
    Mode                := PRG_04_Modes.instModes.Mode,
    SyncEnable          := PRG_04_Modes.instModes.SyncEnable,
    JoystickOnline      := PRG_01_Diagnostics.instDiagCanOpen.Joystick.Online,
    JoystickOperational := PRG_01_Diagnostics.instDiagCanOpen.Joystick.Operational,
    EncoderAvailable    := PRG_02_Encoders.instEncoderAbsM2.EncoderAvailable,
    ThermalFeedback     := NOT PRG_00_Inputs.M2ThermalFeedback,
    BrakeThermalFeedback := NOT PRG_00_Inputs.BrakeThermalFeedback, // 🆕 REX 2026-07-08 — commun M1/M2/M3
    SlackCableDetected  := NOT PRG_00_Inputs.SlackCableSwitch,
    PhaseRotationOk     := PRG_00_Inputs.PhaseRotationOk,
    TopPositionSensor   := PRG_00_Inputs.TopPositionSensor,
    InReferencingMode   := PRG_02_Encoders.instHomingM2.Busy,
    CablePosM           := PRG_02_Encoders.instEncoderScaleM2.CablePosM,
    CableLimitDescentM  := GVL_PERSISTENT.CableLimitDescentM2_M,
    Direction           := PRG_06_WinchControl.M2_Direction_Active,
    Homed               := PRG_02_Encoders.instHomingM2.Homed,
    HomingSuspect       := PRG_02_Encoders.instHomingM2.HomingSuspect,
    TopLimitM           := GVL_PERSISTENT.HomingTargetM2_M,
    // 🔧 REX 2026-07-07 — Méca A/B (voir FB_Safety_Winch bandeau en-tête) — Méca C NON applicable
    // à M2 (c'est M2 qui bouge pendant le grappin, GrappinHoldStillActive reste FALSE)
    FwdRevSpeedFeedbackOff := PRG_00_Inputs.M2FwdRevSpeedFeedbackOff,
    BrakeFeedback          := PRG_00_Inputs.M2BrakeFeedback,
    // 🔧 REX 2026-07-15 (7) : idem M1 (voir bandeau instSafetyWinchM1 ci-dessus).
    JoystickYNeutral       := (ABS(PRG_01_Diagnostics.FB_Joystick_0.AxisCmdY.SpeedRef) < 0.1)
                              AND NOT GVL_IHM.IHM_MANU.M2_RelayFwd AND NOT GVL_IHM.IHM_MANU.M2_RelayRev
                              AND NOT GVL_IHM.IHM_MANU.M1_M2_RelayFwd AND NOT GVL_IHM.IHM_MANU.M1_M2_RelayRev,
    GrappinHoldStillActive := FALSE,
    // 🔧 REX 2026-07-08 (5) : BUG CORRIGÉ — oublié côté M2 lors de l'ajout initial Méca E.
    // ExpectedOtherWinchPosM valait 0.0 par défaut (non câblé) → Méca E comparait CablePosM2
    // à 0 au lieu de M1, déclenchement permanent dès que M2 > CriticalSyncToleranceM (2.0m)
    // du zéro codeur. M1 corrigé de l'offset grappin actif, ramené dans le référentiel M2.
    ExpectedOtherWinchPosM := PRG_02_Encoders.instEncoderScaleM1.CablePosM + PRG_06_WinchControl.instGrappin.ActiveOffsetM,
    GrappinBusy            := PRG_06_WinchControl.instGrappin.Busy,
    CriticalSyncToleranceM := GVL_PERSISTENT.WinchCriticalSyncTolerance_M,
    OtherWinchInhibited    := PRG_04_Modes.instModes.InhibitM1 // 🆕 REX 2026-07-08 (7)
);

// 3. Sécurité Chariot M3
instSafetyChariotM3(
    Enable              := NOT PRG_10_Outputs.ManuActive OR NOT GVL_Simulation.SimulationModeActive OR GVL_Simulation.VariateurM3_IsReal OR GVL_Simulation.ContactorFeedbackM3_IsReal OR GVL_Simulation.ChariotPosition_IsReal, // 🆕 REX 2026-07-14 : ManuActive (Conditional Bypass Doctrine)
    Reset               := PRG_09_Supervision.FaultMachineReset_IHM,
    EmergencyStopOk     := PRG_00_Inputs.EmergencyStopOk,
    Mode                := PRG_04_Modes.instModes.Mode,
    JoystickOnline      := PRG_01_Diagnostics.instDiagCanOpen.Joystick.Online,
    JoystickOperational := PRG_01_Diagnostics.instDiagCanOpen.Joystick.Operational,
    PhaseRotationOk     := PRG_00_Inputs.PhaseRotationOk,
    BrakeThermalFeedback := NOT PRG_00_Inputs.BrakeThermalFeedback, // 🆕 REX 2026-07-08 — commun M1/M2/M3
    DriveOnline         := PRG_01_Diagnostics.instDiagEthercat.Variateur.Online,
    DriveOperational    := PRG_01_Diagnostics.instDiagEthercat.Variateur.Operational,
    DriveStatusWord     := PRG_00_Inputs.M3_StatusWord_Filtered,
    DriveActualFreqHz   := UINT_TO_REAL(PRG_00_Inputs.M3_ActualFrequencyHz_Filtered) / 100.0,
    BrakeFeedback       := PRG_00_Inputs.M3BrakeFeedback,
    BrakeCmd            := PRG_07_ChariotControl.instChariotM3.BrakeCmd,
    Direction           := PRG_07_ChariotControl.M3_Direction_Active,
    LimitSwitchFwd      := PRG_00_Inputs.ChariotPosTremie,
    LimitSwitchRev      := PRG_00_Inputs.ChariotPosFosse1
);

(* ---- PRG_04_Modes.st ---- *)
(* ═══════════════════════════════════════════════════════════════
   🎚️ PRG_04_Modes — Gestion et Arbitrage du Mode Machine
   ───────────────────────────────────────────────────────────────
   ⚙️ Exécuté par la tâche PLC en position 4.
   ═══════════════════════════════════════════════════════════════ *)

PROGRAM PRG_04_Modes
VAR
    instModes : FB_Modes; // Arbitrage du mode machine (DISABLE, MAINT, SEMI_AUTO, etc.)
    PrevInhibitM1 : BOOL; // 🆕 Mémoire d'état M1
    PrevInhibitM2 : BOOL; // 🆕 Mémoire d'état M2
END_VAR

// === IMPLEMENTATION (corps du PROGRAM PRG_04_Modes) ===

// 🆕 Exclusion mutuelle des inhibitions de treuils (soit M1, soit M2, jamais les deux)
IF GVL_IHM.WinchM1.CmdInhibit AND GVL_IHM.WinchM2.CmdInhibit THEN
    // Si M1 était déjà activé, on rejette la demande sur M2 (M2 retombe à FALSE)
    IF PrevInhibitM1 THEN
        GVL_IHM.WinchM2.CmdInhibit := FALSE;
    // Si M2 était déjà activé, on rejette la demande sur M1 (M1 retombe à FALSE)
    ELSIF PrevInhibitM2 THEN
        GVL_IHM.WinchM1.CmdInhibit := FALSE;
    ELSE
        // repli de sécurité si les deux s'activent de façon synchrone sans transition
        GVL_IHM.WinchM1.CmdInhibit := FALSE;
        GVL_IHM.WinchM2.CmdInhibit := FALSE;
    END_IF;
END_IF;

PrevInhibitM1 := GVL_IHM.WinchM1.CmdInhibit;
PrevInhibitM2 := GVL_IHM.WinchM2.CmdInhibit;

// 🆕 Si l'un des treuils est inhibé, synchro impossible par nature -> reset case IHM à TRUE
// (🔧 REX 2026-07-08 : polarité inversée, TRUE = état neutre "synchro voulue")
IF GVL_IHM.WinchM1.CmdInhibit OR GVL_IHM.WinchM2.CmdInhibit THEN
    GVL_IHM.Sync.SyncEnableRequest := TRUE;
END_IF;

instModes(
    Enable              := TRUE,
    Reset               := GVL_IHM.Modes.ModeReset,  // 🔧 REX 2026-07-07 : dédié, jamais mélangé au reset défauts général
    EmergencyStopOk     := PRG_00_Inputs.EmergencyStopOk,
    ModeRequest         := GVL_Modes_Stub.ModeRequest_IHM,      // 🖥️ Sélecteur IHM
    SyncEnableRequest   := GVL_Modes_Stub.SyncEnableRequest_IHM,
    InhibitM1Request    := GVL_IHM.WinchM1.CmdInhibit, // 🆕 REX 2026-07-08 : IHM réelle, pas GVL_Modes_Stub
    InhibitM2Request    := GVL_IHM.WinchM2.CmdInhibit, // 🆕 REX 2026-07-08 : IHM réelle, pas GVL_Modes_Stub
    HomingApproachEnableRequest := GVL_IHM.Common.HomingApproachEnableRequest, // 🆕 REX 2026-07-08 (2)
    EncoderFaultPresent := PRG_02_Encoders.EncoderFaultPresent,   // 1 cycle de retard (reçu de PRG_02_Encoders)
    JoystickWinchSelectRequest := GVL_IHM.IHM_MANU.JoystickWinchSelect // 🆕 TASK-0001
);

(* ---- PRG_05_Cycle.st ---- *)
(* ═══════════════════════════════════════════════════════════════
   🔄 PRG_05_Cycle — Séquenceur du Cycle Automatique / Semi-Auto (Grafcet)
   ───────────────────────────────────────────────────────────────
   ⚙️ Exécuté par la tâche PLC en position 5.
   ✅ Gère la machine d'état principale de dragage (FB_Cycle).
   ═══════════════════════════════════════════════════════════════ *)

PROGRAM PRG_05_Cycle
VAR
    // Instance du séquenceur automatique
    instCycle           : FB_Cycle;

    // Commandes issues de la supervision (IHM)
    CmdStartCycle_IHM   : BOOL;         // Lancement cycle automatique
    CmdPauseCycle_IHM   : BOOL;         // Pause cycle automatique
    CmdAbortCycle_IHM   : BOOL;         // Abandon / arrêt cycle automatique
    CmdResetCycle_IHM   : BOOL;         // 🔧 REX 2026-07-07 : reset dédié FB_Cycle, jamais mélangé au reset défauts général

    // Paramètres cibles réglés par l'opérateur
    TargetDepthM        : REAL := -12.5; // Profondeur de dragage cible (mètres, négative)
    TargetOffsetM       : REAL := 1.5;  // Décalage cible de fermeture du grappin (mètres)
END_VAR

// === IMPLEMENTATION (corps du PROGRAM PRG_05_Cycle) ===

// Appel du séquenceur de cycle principal avec tous ses raccordements
instCycle(
    Enable              := (PRG_04_Modes.instModes.Mode = E_Mode.SEMI_AUTO) AND NOT PRG_10_Outputs.ManuActive,
    Reset               := CmdResetCycle_IHM,
    EmergencyStopOk     := PRG_00_Inputs.EmergencyStopOk,

    StartCycle          := CmdStartCycle_IHM,
    PauseCycle          := CmdPauseCycle_IHM,
    AbortCycle          := CmdAbortCycle_IHM,

    TargetDepthM        := TargetDepthM,
    TargetOffsetM       := TargetOffsetM,
    SelectedTargetNum_IHM := GVL_IHM.ChariotM3.SelectedTargetNum,

    // Capteur fond touché détecté par le mou de câble physique (sécurité positive)
    BottomTouched       := NOT PRG_00_Inputs.SlackCableSwitch,
    M1_CablePosM        := PRG_02_Encoders.instEncoderScaleM1.CablePosM,
    M2_CablePosM        := PRG_02_Encoders.instEncoderScaleM2.CablePosM,

    // Position chariot
    Chariot_At_Fosse1   := PRG_00_Inputs.ChariotPosFosse1,
    Chariot_At_Fosse2   := PRG_00_Inputs.ChariotPosFosse2,
    Chariot_At_Maintenance := PRG_00_Inputs.ChariotPosMaintenance,
    Chariot_At_Tremie   := PRG_00_Inputs.ChariotPosTremie,
    Chariot_Busy        := PRG_07_ChariotControl.instChariotM3.Busy,
    Chariot_Done        := PRG_07_ChariotControl.instChariotM3.Done,

    // Mouvements mâchoires grappin (gérés par instGrappin)
    Grappin_Busy        := PRG_06_WinchControl.instGrappin.Busy,
    Grappin_Done        := PRG_06_WinchControl.instGrappin.Done,
    Grappin_IsOpen      := GVL_PERSISTENT.GrappinState.IsOpen,
    Grappin_IsClosed    := GVL_PERSISTENT.GrappinState.IsClosed
);

(* ---- PRG_06_WinchControl.st ---- *)
(* ═══════════════════════════════════════════════════════════════
   🪝 PRG_06_WinchControl — Commande des Treuils M1/M2, Synchro et Grappin
   ───────────────────────────────────────────────────────────────
   ⚙️ Exécuté par la tâche PLC en position 6.
   ✅ Arbitre entre les commandes Manuelles (Joystick) et Automatiques (PRG_05_Cycle).
   ═══════════════════════════════════════════════════════════════ *)

PROGRAM PRG_06_WinchControl
VAR
    // Stubs
    StubMachineEnableN1 : BOOL := TRUE;

    // Instances
    instWinchSync : FB_WinchSync;
    instGrappin   : FB_Grappin;
    instWinchM1   : FB_Winch;
    instWinchM2   : FB_Winch;

    // Variables de commande M1 après arbitrage Manuel/Auto
    M1_StartStop_Active     : BOOL;
    M1_Direction_Active     : INT;
    M1_SpeedRef_Active      : REAL;

    // Variables de commande M2 après arbitrage Grappin/Manuel/Auto
    M2_StartStop_Active     : BOOL;
    M2_Direction_Active     : INT;
    M2_SpeedRef_Active      : REAL;
    M2_SpeedStepTableActive : ST_SpeedStepTable;

    // Bornage et limites
    BottomLimitM1_Active    : REAL;
    BottomLimitM2_Active    : REAL;
    ForbidDescentM1_Active  : BOOL;
    ForbidDescentM2_Active  : BOOL;
    // 🆕 REX 2026-07-15 (8) — miroir IHM dédié CableLimitAscentM1/2_M (demande utilisateur, symétrique
    // à CableLimitDescentReached) : indique PRÉCISÉMENT que la nouvelle limite haute d'exploitation
    // normale est atteinte (hors capteur physique bit5, hors Homing) — voir §5 plus bas.
    CableLimitAscentM1Reached : BOOL;
    CableLimitAscentM2Reached : BOOL;

    // 🔧 REX 2026-07-07 : couplage croisé M1/M2 des arrêts, UNIQUEMENT si SyncActive (mouvement
    // coherent voulu). Hors synchro (Grappin.Busy ou SyncEnable=FALSE MAINT_N2) : chaque treuil réagit
    // à SA PROPRE limite/défaut uniquement — commande indépendante voulue dans ce cas.
    SafeStopM1_Raw          : BOOL;
    SafeStopM2_Raw          : BOOL;
    SafeStopM1_Active       : BOOL;
    SafeStopM2_Active       : BOOL;
    ForbidDescentM1_Raw     : BOOL;
    ForbidDescentM2_Raw     : BOOL;
    ForbidAscentM1_Raw      : BOOL;
    ForbidAscentM2_Raw      : BOOL;
    ForbidAscentM1_Active   : BOOL;
    ForbidAscentM2_Active   : BOOL;

    // 🆕 REX 2026-07-08 : voir §2bis — coupure immédiate M1/M2 au même scan que la fin du cycle
    // grappin (contrairement au désarmement homme-mort côté FB_Joystick, qui a 1 scan de retard
    // structurel — PRG_01 s'exécute avant PRG_06). Corrige un bref "blip" de commande (RelayFwd/Rev
    // + BrakeCmd clignotant) observé sur M1 à l'arrivée en position grappin.
    GrappinBusyFallEdge     : F_TRIG;

    // 🆕 REX 2026-07-08 (4) : instWinchSync appelé APRÈS l'arbitrage M1/M2 (§3, plus bas) — lu ici
    // avec 1 scan de retard (~10ms), négligeable vu que DeltaPosM évolue progressivement, pas
    // par à-coup (même raisonnement que M1_Busy/M2_Busy sur instGrappin, voir §0).
    SyncMinorDeviation      : BOOL;
    SyncMinorDeviationBlocksUp   : BOOL;   // 🆕 REX 2026-07-08 (5) : bit0 latché ET écart actuel aggravé par la montée
    SyncMinorDeviationBlocksDown : BOOL;   // 🆕 REX 2026-07-08 (5) : bit0 latché ET écart actuel aggravé par la descente
    M2_LimitShift                : REAL;   // 🆕 REX 2026-07-08 : décalage dynamique de la butée haute de M2

    // 🆕 REX 2026-07-15 (3) — demande utilisateur : les fins de course virtuelles grappin
    // (FdcGrappinOpen/CloseActive) doivent bloquer le mouvement AUSSI en pilotage COUPLÉ IHM_MANU
    // (M1+M2 simultané), pas seulement en pilotage individuel M2 — sinon un opérateur qui pousse le
    // couplage alors que le grappin est déjà en butée virtuelle n'est protégé que par la butée
    // mécanique passive. Masque calculé UNE FOIS ici, consommé par M1 ET M2 (§1/§2 ci-dessous) pour
    // que les deux treuils s'arrêtent ENSEMBLE (pas de désynchro M1/M2 en cas de blocage partiel).
    CoupledFwdGrappinOk          : BOOL;   // Couplage montée autorisé (pas de butée fermeture grappin)
    CoupledRevGrappinOk          : BOOL;   // Couplage descente autorisé (pas de butée ouverture grappin)

    // 🆕 REX 2026-07-15 (9) — plafond palier IHM_MANU "essais progressifs" (demande utilisateur,
    // TEMPORAIRE tant que les vitesses définitives ne sont pas figées, à retirer ensuite) : commun
    // aux 2 treuils (GVL_IHM.IHM_MANU.WinchMaxStepFwd/Rev, structure figée, un seul réglage pour M1
    // ET M2). Actif UNIQUEMENT si ManuActive — Auto garde son comportement inchangé (5 en montée,
    // WinchMaxStepDescente en descente). En Manu, le plafond descente est le MIN avec
    // WinchMaxStepDescente (jamais moins protecteur qu'Auto, juste potentiellement plus prudent).
    ManuMaxStepFwd            : INT;
    ManuMaxStepRev            : INT;
    EffectiveMaxStepAscent    : INT;
    EffectiveMaxStepDescente  : INT;
END_VAR

// === IMPLEMENTATION (corps du PROGRAM PRG_06_WinchControl) ===

// ── 0. COMMANDE DU GRAPPIN (Séquence lente) ─────────────────────────────
// 🔧 REX 2026-07-08 : appelé EN PREMIER (avant l'arbitrage M1/M2 ci-dessous) — audit sécurité :
// l'ancien ordre (Grappin appelé après l'arbitrage) faisait que M1_StartStop_Active lisait
// instGrappin.Busy du scan PRÉCÉDENT, créant une fenêtre d'1 scan où M1 pouvait recevoir une
// commande manuelle au moment exact où le grappin démarre. instGrappin.M1_Busy/M2_Busy (ci-dessous)
// lisent en retour instWinchM1/M2.Busy du scan précédent (ces FB sont appelés plus loin, §6/§7) —
// acceptable : ça ne retarde que l'ACCEPTATION d'une nouvelle demande de ~1 scan (10ms), sans
// aucun impact sécurité (contrairement au cas inverse, qui pouvait faire bouger M1 pendant Busy).
instGrappin(
    Enable              := NOT PRG_04_Modes.instModes.InhibitM2
                           AND PRG_02_Encoders.instEncoderAbsM1.EncoderAvailable
                           AND PRG_02_Encoders.instEncoderAbsM2.EncoderAvailable, // 🆕 Sécurisé : nécessite les deux codeurs valides et M2 non-inhibé
    Reset               := PRG_09_Supervision.FaultMachineReset_IHM,
    EmergencyStopOk     := PRG_00_Inputs.EmergencyStopOk,
    Mode                := PRG_04_Modes.instModes.Mode,
    CmdOpen_IHM         := GVL_IHM.Grappin.CmdOpen OR PRG_05_Cycle.instCycle.CmdGrappin_Open,
    CmdClose_IHM        := GVL_IHM.Grappin.CmdClose OR PRG_05_Cycle.instCycle.CmdGrappin_Close,
    JoystickY_StartStop := PRG_01_Diagnostics.FB_Joystick_0.AxisCmdY.StartStop,
    JoystickY_Direction := PRG_01_Diagnostics.FB_Joystick_0.AxisCmdY.Direction,
    CablePosM1          := PRG_02_Encoders.instEncoderScaleM1.CablePosM,
    CablePosM2          := PRG_02_Encoders.instEncoderScaleM2.CablePosM,
    HomedM1             := PRG_02_Encoders.instHomingM1.Homed,
    HomedM2             := PRG_02_Encoders.instHomingM2.Homed,
    M1_Busy             := instWinchM1.Busy,   // 🆕 REX 2026-07-08
    M2_Busy             := instWinchM2.Busy,   // 🆕 REX 2026-07-08
    ConfirmOpenPosition := GVL_IHM.Grappin.CmdConfirmOpenPosition, // 🆕 REX 2026-07-08 — bouton IHM référencement grappin ouvert
    ConfirmClosePosition:= GVL_IHM.Grappin.CmdConfirmClosePosition, // 🆕 REX 2026-07-08 — bouton IHM référencement grappin fermé
    Config              := GVL_PERSISTENT.GrappinConfig,
    TimeoutDuration     := GVL_IHM.Grappin.TimeoutDuration,
    GrappinState        := GVL_PERSISTENT.GrappinState,
    InhibitM1           := PRG_04_Modes.instModes.InhibitM1, // 🆕 REX 2026-07-08
    InhibitM2           := PRG_04_Modes.instModes.InhibitM2  // 🆕 REX 2026-07-08
);

// 🆕 REX 2026-07-08 (4) — Concept 1 (écart synchro mineur) : bit0 seul (écart position, hors
// incohérence commande bit1) ne fait plus de SafeStop (fast) — bloque StartStop → rampe de décél
// NORMALE. Recalage : voir SyncEnable=FALSE (MAINT_N2), procédure déjà existante (mou de câble).
SyncMinorDeviation := (instWinchSync.ErrorId AND 16#0001) <> 16#0000;

// 🔧 REX 2026-07-08 (5) — audit sécurité : ne bloque plus StartStop dans les 2 sens (déblocage
// impossible sans Reset+MAINT_N2, régression terrain constatée, écart mécanique transitoire
// normal à l'arrêt). SignedDeltaPosM > 0 = M1 plus "haut" que M2 : la montée (Direction=+1)
// aggrave cet écart, la descente (-1) le réduit — et inversement si < 0. Seul le sens aggravant
// reste bloqué ; Méca E (FB_Safety_Winch, écart critique 2.0m) et bit1 (incohérence commande)
// restent le filet réel si l'écart continue de dériver malgré cette autorisation directionnelle.
// 🆕 REX 2026-07-08 (6) : gate global SyncSoftStopEnable — FALSE (défaut) = ces 2 sorties
// restent FALSE en permanence (bit0 déjà géré en SafeStop fast classique ci-dessus, §5bis) ;
// TRUE = active le blocage directionnel (nouvelle fonctionnalité, opt-in).
SyncMinorDeviationBlocksUp   := GVL_PERSISTENT.SyncSoftStopEnable AND SyncMinorDeviation AND (instWinchSync.SignedDeltaPosM > 0.0);
SyncMinorDeviationBlocksDown := GVL_PERSISTENT.SyncSoftStopEnable AND SyncMinorDeviation AND (instWinchSync.SignedDeltaPosM < 0.0);

// 🆕 REX 2026-07-15 (3) — voir déclaration VAR ci-dessus : couplé masqué par les mêmes fins de
// course grappin que l'individuel M2, appliqué à M1 ET M2 (§1/§2) pour arrêter les DEUX treuils
// ensemble plutôt que de désynchroniser M1/M2 en ne bloquant que la moitié du couplage.
CoupledFwdGrappinOk := NOT GVL_IHM.IHM_MANU.FdcGrappinCloseActive;
CoupledRevGrappinOk := NOT GVL_IHM.IHM_MANU.FdcGrappinOpenActive;

// 🆕 REX 2026-07-15 (9) — plafond palier IHM_MANU "essais progressifs" (voir déclaration VAR
// ci-dessus). Bornage identique à l'ex-logique PRG_10_Outputs retirée lors du passage sur FB_Winch.
ManuMaxStepFwd := GVL_IHM.IHM_MANU.WinchMaxStepFwd;
IF (ManuMaxStepFwd < 1) OR (ManuMaxStepFwd > 5) THEN
    ManuMaxStepFwd := 5; // Pleine vitesse par défaut si non initialisé/invalide
END_IF;
ManuMaxStepRev := GVL_IHM.IHM_MANU.WinchMaxStepRev;
IF (ManuMaxStepRev < 1) OR (ManuMaxStepRev > 5) THEN
    ManuMaxStepRev := 2; // Palier 2 max par défaut en descente (conforme AF) si non initialisé/invalide
END_IF;
EffectiveMaxStepAscent   := SEL(PRG_10_Outputs.ManuActive, 5, ManuMaxStepFwd);
EffectiveMaxStepDescente := SEL(PRG_10_Outputs.ManuActive, GVL_PERSISTENT.WinchMaxStepDescente, MIN(GVL_PERSISTENT.WinchMaxStepDescente, ManuMaxStepRev));

// ── 1. ARBITRAGE DES CONSIGNES M1 (Joystick vs Cycle Automatique) ────────
IF PRG_04_Modes.instModes.Mode = E_Mode.SEMI_AUTO THEN
    // 🔧 REX 2026-07-08 (7) — review : gate directionnel absent de cette branche (bug trouvé en
    // review code), le cycle auto pouvait aggraver un écart mineur sans aucune protection quand
    // SyncSoftStopEnable=TRUE. Ajouté ici, symétrique à la branche manuelle ci-dessous.
    M1_Direction_Active := PRG_05_Cycle.instCycle.CmdWinchM1_Direction;
    M1_StartStop_Active := PRG_05_Cycle.instCycle.CmdWinchM1_StartStop
                            AND NOT ((SyncMinorDeviationBlocksUp   AND (M1_Direction_Active = 1))
                                 OR  (SyncMinorDeviationBlocksDown AND (M1_Direction_Active = -1)));
    M1_SpeedRef_Active  := PRG_05_Cycle.instCycle.CmdWinchM1_SpeedPct;
ELSIF PRG_10_Outputs.ManuActive THEN
    // 🆕 REX 2026-07-15 (2) — IHM_MANU pilote désormais M1 via FB_Winch (au lieu de l'ex-bypass
    // direct dans PRG_10_Outputs) : récupère gratuitement la rampe accel/décel + le ralentissement
    // en zone d'approche de bordure + le maintien du relais pendant la décél (mêmes paramètres
    // persistants qu'en Auto, voir instWinchM1 plus bas §6). Demande (boutons IHM ou joystick, déjà
    // arbitrée par PRG_10_Outputs : M1Fwd_Demand/M1Rev_Demand/CoupledFwd_Demand/CoupledRev_Demand)
    // lue avec 1 scan de retard (~10ms, PRG_10 position 10 > PRG_06 position 6) — même principe
    // déjà accepté ailleurs dans ce fichier (Grappin.Busy, SyncMinorDeviation).
    // 🔧 REX 2026-07-15 (5) — trouvé en revue croisée (agent Haiku + relecture manuelle) : M1
    // INDIVIDUEL (bouton M1_RelayFwd/Rev, indépendant de M2) n'était masqué par AUCUNE butée
    // grappin — delta = CablePosM1 - CablePosM2, donc bouger M1 seul aggrave la MÊME sur-contrainte
    // mécanique que le couplé (déjà corrigé ci-dessous) : M1 Fwd augmente le delta (aggrave
    // FdcGrappinOpenActive, delta déjà >= 0) ; M1 Rev diminue le delta (aggrave
    // FdcGrappinCloseActive, delta déjà <= -10). Sens INVERSÉ par rapport à M2 (M2Fwd↔Close,
    // M2Rev↔Open) car M1 et M2 ont un effet opposé sur le même delta. Couplé masqué par
    // CoupledFwdGrappinOk/CoupledRevGrappinOk (REX 2026-07-15 (3)) — M1 s'arrête EN MÊME TEMPS que
    // M2 si le couplage OU son propre individuel violerait une butée grappin.
    IF (PRG_10_Outputs.M1Fwd_Demand AND NOT GVL_IHM.IHM_MANU.FdcGrappinOpenActive) OR (PRG_10_Outputs.CoupledFwd_Demand AND CoupledFwdGrappinOk) THEN
        M1_Direction_Active := 1;
    ELSIF (PRG_10_Outputs.M1Rev_Demand AND NOT GVL_IHM.IHM_MANU.FdcGrappinCloseActive) OR (PRG_10_Outputs.CoupledRev_Demand AND CoupledRevGrappinOk) THEN
        M1_Direction_Active := -1;
    ELSE
        M1_Direction_Active := 0;
    END_IF;
    M1_StartStop_Active := (M1_Direction_Active <> 0);
    // 🎯 Joystick = vitesse proportionnelle à la déflexion (comme en Auto) ; boutons HMI = cible 100%
    // (FB_Winch rampe déjà en interne, plus besoin de la rampe HMI locale ex-PRG_10_Outputs).
    M1_SpeedRef_Active  := SEL(GVL_IHM.IHM_MANU.JoystickSelect, 100.0, ABS(PRG_01_Diagnostics.FB_Joystick_0.AxisCmdY.SpeedRef));
ELSE
    // 🔧 REX 2026-07-08 : + AND DeadmanArmed — NOT Busy seul insuffisant (rampe joystick met du
    // temps à redescendre à 0 après désarmement homme-mort ⇒ StartStop reste TRUE le temps de la
    // décél, M1 bougeait/frein décollait à la fin d'un cycle grappin). DeadmanArmed reste FALSE
    // en continu jusqu'au repassage neutre + réappui, sans dépendre du temps de rampe.
    // 🔧 REX 2026-07-08 (5) : Direction assignée AVANT StartStop (nécessaire pour le gate directionnel ci-dessous).
    M1_Direction_Active := PRG_01_Diagnostics.FB_Joystick_0.AxisCmdY.Direction;
    M1_StartStop_Active := PRG_01_Diagnostics.FB_Joystick_0.AxisCmdY.StartStop AND NOT instGrappin.Busy
                            AND PRG_01_Diagnostics.FB_Joystick_0.DeadmanArmed
                            AND NOT ((SyncMinorDeviationBlocksUp   AND (M1_Direction_Active = 1))
                                 OR  (SyncMinorDeviationBlocksDown AND (M1_Direction_Active = -1))); // 🔧 REX 2026-07-08 (5)
    M1_SpeedRef_Active  := PRG_01_Diagnostics.FB_Joystick_0.AxisCmdY.SpeedRef;
END_IF;

// ── 2. ARBITRAGE DES CONSIGNES M2 (Grappin vs Cycle Automatique vs Joystick) ──
IF instGrappin.Busy THEN
    M2_StartStop_Active := instGrappin.M2_StartStop;
    M2_Direction_Active := instGrappin.M2_Direction;
    M2_SpeedRef_Active  := 15.0; // Vitesse lente forcée pour fermeture grappin
ELSE
    IF PRG_04_Modes.instModes.Mode = E_Mode.SEMI_AUTO THEN
        // 🔧 REX 2026-07-08 (7) — review : gate directionnel absent de cette branche, ajouté
        // symétrique à la branche manuelle ci-dessous (signe M2, voir note ci-dessous).
        M2_Direction_Active := PRG_05_Cycle.instCycle.CmdWinchM2_Direction;
        M2_StartStop_Active := PRG_05_Cycle.instCycle.CmdWinchM2_StartStop
                                AND NOT ((SyncMinorDeviationBlocksUp   AND (M2_Direction_Active = -1))
                                     OR  (SyncMinorDeviationBlocksDown AND (M2_Direction_Active = 1)));
        M2_SpeedRef_Active  := PRG_05_Cycle.instCycle.CmdWinchM2_SpeedPct;
    ELSIF PRG_10_Outputs.ManuActive THEN
        // 🔧 REX 2026-07-15 (3) — idem M1 (voir §1) : Fins de course grappin (FdcGrappin) appliquées
        // au pilotage INDIVIDUEL **ET** COUPLÉ de M2 désormais (demande utilisateur — "que ce soit
        // couplé ou pas couplé, il faut rester dans les butées"). Ex-comportement (couplé non
        // masqué) retiré : c'était une incohérence, pas un choix voulu.
        IF (PRG_10_Outputs.M2Fwd_Demand AND NOT GVL_IHM.IHM_MANU.FdcGrappinCloseActive) OR (PRG_10_Outputs.CoupledFwd_Demand AND CoupledFwdGrappinOk) THEN
            M2_Direction_Active := 1;
        ELSIF (PRG_10_Outputs.M2Rev_Demand AND NOT GVL_IHM.IHM_MANU.FdcGrappinOpenActive) OR (PRG_10_Outputs.CoupledRev_Demand AND CoupledRevGrappinOk) THEN
            M2_Direction_Active := -1;
        ELSE
            M2_Direction_Active := 0;
        END_IF;
        M2_StartStop_Active := (M2_Direction_Active <> 0);
        M2_SpeedRef_Active  := SEL(GVL_IHM.IHM_MANU.JoystickSelect, 100.0, ABS(PRG_01_Diagnostics.FB_Joystick_0.AxisCmdY.SpeedRef));
    ELSE
        // 🔧 REX 2026-07-08 : + AND DeadmanArmed, même raison que M1 ci-dessus
        // 🔧 REX 2026-07-08 (5) : Direction assignée AVANT StartStop (gate directionnel)
        // 🐛 REX 2026-07-08 (7) — BUG CORRIGÉ (review code) : signe inversé pour M2. SignedDeltaPosM
        // (référentiel M1 : CablePosM1-CablePosM2+Offset) > 0 signifie M1 en avance — pour RATTRAPER,
        // M2 doit MONTER (+1), pas descendre. Donc BlocksUp (écart M1-en-avance) doit bloquer côté M2
        // le sens qui AGGRAVE, c-à-d Direction=-1 (descendre, M2 prend encore plus de retard) — PAS
        // Direction=+1 (monter, qui RATTRAPE). Symétrique inversé par rapport à M1 (qui utilise +1/-1
        // directement car SignedDeltaPosM est déjà dans SON référentiel).
        M2_Direction_Active := PRG_01_Diagnostics.FB_Joystick_0.AxisCmdY.Direction;
        M2_StartStop_Active := PRG_01_Diagnostics.FB_Joystick_0.AxisCmdY.StartStop
                                AND PRG_01_Diagnostics.FB_Joystick_0.DeadmanArmed
                                AND NOT ((SyncMinorDeviationBlocksUp   AND (M2_Direction_Active = -1))
                                     OR  (SyncMinorDeviationBlocksDown AND (M2_Direction_Active = 1))); // 🔧 REX 2026-07-08 (7)
        M2_SpeedRef_Active  := PRG_01_Diagnostics.FB_Joystick_0.AxisCmdY.SpeedRef;
    END_IF;
END_IF;

// ── 2bis. COUPURE IMMÉDIATE M1/M2 AU SCAN EXACT DE FIN DE CYCLE GRAPPIN ─────
// 🆕 REX 2026-07-08 : instGrappin est appelé en premier (§0), donc son Busy est frais dans CE scan
// (voir §1/§2 ci-dessus) — mais AxisCmdY.StartStop/Direction viennent de FB_Joystick_0 (PRG_01),
// calculé AVANT ce scan de PRG_06. Le désarmement homme-mort sur front descendant de Grappin.Busy
// (FB_Joystick §4ter-ter) ne prend donc effet qu'au scan SUIVANT (~10ms de retard structurel). Si
// l'opérateur tient encore le manche poussé au moment exact où le grappin termine, M1 ET M2
// recevaient pendant ce scan la commande manche brute (RelayFwd/Rev + BrakeCmd qui s'engage puis se
// coupe aussitôt = "clignotement" du frein, constaté sur site). On force ici l'arrêt immédiat,
// sans attendre le désarmement (qui reste nécessaire pour la suite : repassage au neutre exigé).
GrappinBusyFallEdge(CLK := instGrappin.Busy);
IF GrappinBusyFallEdge.Q THEN
    M1_StartStop_Active := FALSE;
    M2_StartStop_Active := FALSE;
END_IF;

// ── 3. SURVEILLANCE ÉCART DE SYNCHRONISATION ────────────────────────────
instWinchSync(
    // 🐛 REX 2026-07-08 (7) — BUG CORRIGÉ (retour terrain, simulation) : écart transitoire (~0.27m)
    // constaté UNIQUEMENT à l'approche d'une butée (haute 12m ici), pas pendant le pilotage normal
    // (précision <0.001m confirmée par l'opérateur). Cause : ForbidAscent/ForbidDescent coupent
    // M1/M2 au même scan (couplage croisé), mais leur arrêt PHYSIQUE (rampe de décél, même en
    // simulation) n'est jamais parfaitement simultané à la position exacte — écart normal et non
    // significatif à ce moment précis, pas une vraie désynchro. Suppression pendant qu'un des deux
    // treuils est en butée (Ascent OU Descent), même principe que la suppression pendant GrappinBusy
    // déjà existante. Lu avec 1 scan de retard (ForbidAscent/DescentMx_Active calculés plus bas dans
    // ce fichier) — acceptable, même raisonnement que SyncMinorDeviation ci-dessous.
    Enable          := PRG_04_Modes.instModes.SyncEnable AND NOT instGrappin.Busy
                        AND NOT PRG_04_Modes.instModes.InhibitM1 AND NOT PRG_04_Modes.instModes.InhibitM2
                        AND NOT (ForbidAscentM1_Active OR ForbidAscentM2_Active
                                 OR ForbidDescentM1_Active OR ForbidDescentM2_Active), // 🆕 REX 2026-07-08 (7)
    Reset           := PRG_09_Supervision.FaultMachineReset_IHM,
    EmergencyStopOk := PRG_00_Inputs.EmergencyStopOk,
    Mode            := PRG_04_Modes.instModes.Mode,
    CablePosM1      := PRG_02_Encoders.instEncoderScaleM1.CablePosM,
    CablePosM2      := PRG_02_Encoders.instEncoderScaleM2.CablePosM,
    HomedM1         := PRG_02_Encoders.instHomingM1.Homed,
    HomedM2         := PRG_02_Encoders.instHomingM2.Homed,
    SyncEnable      := PRG_04_Modes.instModes.SyncEnable,
    SyncToleranceM  := GVL_PERSISTENT.WinchSyncTolerance_M,
    ActiveOffsetM   := instGrappin.ActiveOffsetM,

    RelayFwdM1      := instWinchM1.RelayFwd,
    RelayFwdM2      := instWinchM2.RelayFwd,
    RelayRevM1      := instWinchM1.RelayRev,
    RelayRevM2      := instWinchM2.RelayRev,
    Contactor1_M1   := instWinchM1.Contactor1,
    Contactor1_M2   := instWinchM2.Contactor1,
    Contactor2_M1   := instWinchM1.Contactor2,
    Contactor2_M2   := instWinchM2.Contactor2,
    Contactor3_M1   := instWinchM1.Contactor3,
    Contactor3_M2   := instWinchM2.Contactor3,
    Contactor4_M1   := instWinchM1.Contactor4,
    Contactor4_M2   := instWinchM2.Contactor4
);

// Table active M2 (verrouille TOUS les paliers sur la combinaison réelle du palier 1 si
// vitesse lente requise pour le grappin — REX 2026-07-08 : l'ancienne version mettait
// TOUS les contacteurs à FALSE pour tous les paliers, y compris le palier 1 lui-même, ce qui
// donnait un mouvement à vitesse quasi nulle/insuffisante (résistance rotorique maximale, aucun
// contacteur de vitesse engagé). Le palier 1 réel (`WinchSpeedStepTable.P1Rx`) engage déjà le
// contacteur le plus lent prévu pour un fonctionnement normal — on le duplique sur les 5 paliers
// pour que M2 reste TOUJOURS à cette vitesse pendant le grappin, quelle que soit l'amplitude
// joystick (peu importe le palier sélectionné par l'hystérésis, le résultat est identique).
IF instGrappin.M2_ForceSlowSpeed THEN
    M2_SpeedStepTableActive.P1R1 := GVL_PERSISTENT.WinchSpeedStepTable.P1R1;
    M2_SpeedStepTableActive.P1R2 := GVL_PERSISTENT.WinchSpeedStepTable.P1R2;
    M2_SpeedStepTableActive.P1R3 := GVL_PERSISTENT.WinchSpeedStepTable.P1R3;
    M2_SpeedStepTableActive.P1R4 := GVL_PERSISTENT.WinchSpeedStepTable.P1R4;
    M2_SpeedStepTableActive.P2R1 := GVL_PERSISTENT.WinchSpeedStepTable.P1R1;
    M2_SpeedStepTableActive.P2R2 := GVL_PERSISTENT.WinchSpeedStepTable.P1R2;
    M2_SpeedStepTableActive.P2R3 := GVL_PERSISTENT.WinchSpeedStepTable.P1R3;
    M2_SpeedStepTableActive.P2R4 := GVL_PERSISTENT.WinchSpeedStepTable.P1R4;
    M2_SpeedStepTableActive.P3R1 := GVL_PERSISTENT.WinchSpeedStepTable.P1R1;
    M2_SpeedStepTableActive.P3R2 := GVL_PERSISTENT.WinchSpeedStepTable.P1R2;
    M2_SpeedStepTableActive.P3R3 := GVL_PERSISTENT.WinchSpeedStepTable.P1R3;
    M2_SpeedStepTableActive.P3R4 := GVL_PERSISTENT.WinchSpeedStepTable.P1R4;
    M2_SpeedStepTableActive.P4R1 := GVL_PERSISTENT.WinchSpeedStepTable.P1R1;
    M2_SpeedStepTableActive.P4R2 := GVL_PERSISTENT.WinchSpeedStepTable.P1R2;
    M2_SpeedStepTableActive.P4R3 := GVL_PERSISTENT.WinchSpeedStepTable.P1R3;
    M2_SpeedStepTableActive.P4R4 := GVL_PERSISTENT.WinchSpeedStepTable.P1R4;
    M2_SpeedStepTableActive.P5R1 := GVL_PERSISTENT.WinchSpeedStepTable.P1R1;
    M2_SpeedStepTableActive.P5R2 := GVL_PERSISTENT.WinchSpeedStepTable.P1R2;
    M2_SpeedStepTableActive.P5R3 := GVL_PERSISTENT.WinchSpeedStepTable.P1R3;
    M2_SpeedStepTableActive.P5R4 := GVL_PERSISTENT.WinchSpeedStepTable.P1R4;
    M2_SpeedStepTableActive.StepThreshold_Pct := GVL_PERSISTENT.WinchSpeedStepTable.StepThreshold_Pct;
ELSE
    M2_SpeedStepTableActive := GVL_PERSISTENT.WinchSpeedStepTable;
END_IF;

// ── 5. CALCUL DES LIMITES BASSES ACTIVES ET DU BLOCAGE DE DESCENTE ──────
// 🔧 REX 2026-07-07 : limite légale appliquée sur LimitLegalEnabled SEUL, plus de garde
// Mode=SEMI_AUTO — la limite légale doit stopper la descente dans TOUS les modes dès qu'elle
// est activée (constat terrain : ne s'arrêtait pas en MAINT_N1/N2 alors qu'attendu).
BottomLimitM1_Active := GVL_PERSISTENT.CableLimitDescentM1_M;
IF GVL_PERSISTENT.LimitLegalEnabled THEN
    BottomLimitM1_Active := MAX(BottomLimitM1_Active, GVL_PERSISTENT.LimitLegalDepthMinAllowed);
END_IF;

BottomLimitM2_Active := GVL_PERSISTENT.CableLimitDescentM2_M;
IF GVL_PERSISTENT.LimitLegalEnabled THEN
    BottomLimitM2_Active := MAX(BottomLimitM2_Active, GVL_PERSISTENT.LimitLegalDepthMinAllowed);
END_IF;

// ── 5bis. COUPLAGE CROISÉ M1/M2 — REX 2026-07-07 ────────────────────────
// Hors synchro (Grappin.Busy ou SyncEnable=FALSE N2) : chaque treuil réagit à SA PROPRE limite/
// défaut uniquement (commande indépendante voulue). En synchro (SyncActive, mouvement cohérent
// voulu) : n'importe quel arrêt (SafeStop, limite câble, limite légale, fin de course haut) sur
// UN treuil coupe IMMÉDIATEMENT les deux — pas d'attente du filtre 500ms de FB_WinchSync.
// 🔧 REX 2026-07-07 : instGrappin.M1SlipDetected ajouté à M1 uniquement (Méca C couche 1) — M2
// est déjà arrêté par son propre mécanisme SevereError interne à FB_Grappin, pas besoin ici.
// 🔧 REX 2026-07-08 (4) : instWinchSync.Error (bit0+bit1) → SEUL bit1 (incohérence commande,
// grave) reste ici en SafeStop fast. Bit0 (écart mineur) → arrêt rampe normale via StartStop
// (voir SyncMinorDeviation, §1/§2 plus haut) — Concept 1, ne pas dégrader le comportement voulu.
// 🆕 REX 2026-07-08 (6) : GVL_PERSISTENT.SyncSoftStopEnable=FALSE (défaut) → comportement D'AVANT,
// bit0 réintégré ici en SafeStop fast classique comme n'importe quel autre défaut winch. TRUE →
// bit0 exclu d'ici, géré exclusivement par le gate directionnel StartStop (§1/§2).
SafeStopM1_Raw      := PRG_03_Safety.instSafetyWinchM1.SafeStop
                       OR ((instWinchSync.ErrorId AND 16#0002) <> 16#0000)
                       OR (NOT GVL_PERSISTENT.SyncSoftStopEnable AND ((instWinchSync.ErrorId AND 16#0001) <> 16#0000))
                       OR instGrappin.M1SlipDetected;
SafeStopM2_Raw      := PRG_03_Safety.instSafetyWinchM2.SafeStop
                       OR ((instWinchSync.ErrorId AND 16#0002) <> 16#0000)
                       OR (NOT GVL_PERSISTENT.SyncSoftStopEnable AND ((instWinchSync.ErrorId AND 16#0001) <> 16#0000));

ForbidDescentM1_Raw := PRG_03_Safety.instSafetyWinchM1.ForbidDescent
                       OR (GVL_PERSISTENT.LimitLegalEnabled
                           AND (PRG_02_Encoders.instEncoderScaleM1.CablePosM <= GVL_PERSISTENT.LimitLegalDepthMinAllowed));
ForbidDescentM2_Raw := PRG_03_Safety.instSafetyWinchM2.ForbidDescent
                       OR (GVL_PERSISTENT.LimitLegalEnabled
                           AND (PRG_02_Encoders.instEncoderScaleM2.CablePosM <= GVL_PERSISTENT.LimitLegalDepthMinAllowed));

// 🔧 REX 2026-07-15 (6) — demande utilisateur : arrêt réel encodeur en fonctionnement NORMAL,
// distinct du capteur physique (bit5/Méca D côté FB_Safety_Winch). Seuil = CableLimitAscentMx_M,
// limite ABSOLUE indépendante (même principe que CableLimitDescentM1/2_M côté descente) —
// ex-calcul en MARGE sous HomingTargetMx_M (WinchTopStopMarginM) RETIRÉ : HomingTargetMx_M (12.5m)
// est réservée à l'approche petite vitesse du capteur physique pendant un Homing explicite, PAS
// à l'exploitation normale, qui doit s'arrêter proprement BIEN AVANT (12.0m par défaut) sans
// jamais réveiller le capteur physique (bit5/Méca D traitent son activation hors référencement
// comme une ANOMALIE — roue libre/contacteur collé — pas un fonctionnement normal).
// Même principe que la limite légale de descente ci-dessus (condition LIVE, pas de bit
// ErrorId/Reset dédié) — passe par ForbidAscentMx_Raw pour bénéficier DU MÊME couplage croisé
// M1/M2 que le capteur physique (sinon un treuil qui atteint la limite une fraction de seconde
// avant l'autre crée un écart RelayFwdM1<>RelayFwdM2 qui déclenche à tort le défaut FB_WinchSync
// bit1 "incohérence de commande" — REX terrain 2026-07-08, testé et corrigé).
// Bypass en MAINT_N2 via `HomingApproachEnable` (FB_Modes, même pattern que SyncEnable) :
// nécessite MAINT_N2 ET une case IHM activée consciemment pour dépasser CableLimitAscentMx_M
// et aller chercher le capteur physique en petite vitesse (Homing).
// 🆕 REX 2026-07-15 (8) : flag dédié — miroir IHM (GVL_IHM.WinchM1.CableLimitAscentReached, voir
// PRG_09_Supervision), symétrique à CableLimitDescentReached. Réutilisé ci-dessous dans ForbidAscentM1_Raw.
CableLimitAscentM1Reached := PRG_02_Encoders.instHomingM1.Homed
                             AND NOT PRG_02_Encoders.instHomingM1.HomingSuspect
                             AND (PRG_02_Encoders.instEncoderScaleM1.CablePosM >= GVL_PERSISTENT.CableLimitAscentM1_M)
                             AND NOT PRG_04_Modes.instModes.HomingApproachEnable;

ForbidAscentM1_Raw  := PRG_03_Safety.instSafetyWinchM1.ForbidAscent
                       OR (PRG_02_Encoders.instHomingM1.Homed
                           AND NOT PRG_02_Encoders.instHomingM1.HomingSuspect
                           AND (PRG_02_Encoders.instEncoderScaleM1.CablePosM >= GVL_PERSISTENT.HomingTargetM1_M))
                       OR CableLimitAscentM1Reached;
// 🐛 REX 2026-07-08 (7) — BUG CORRIGÉ (retour terrain) / REX 2026-07-08 (2) :
// La butée haute de M2 n'est décalée de l'OffsetCloseM QUE si le grappin est fermé (IsClosed)
// ou en cours de fermeture (CloseReq). Sinon (grappin ouvert/en cours d'ouverture), M2 doit
// s'arrêter à la butée normale (CableLimitAscentM2_M) pour s'arrêter proprement en même temps que M1.
M2_LimitShift := SEL(GVL_PERSISTENT.GrappinState.IsClosed OR instGrappin.CloseReq, 0.0, GVL_PERSISTENT.GrappinConfig.OffsetCloseM);

// 🆕 REX 2026-07-15 (8) : idem M1 (voir ci-dessus).
CableLimitAscentM2Reached := PRG_02_Encoders.instHomingM2.Homed
                             AND NOT PRG_02_Encoders.instHomingM2.HomingSuspect
                             AND (PRG_02_Encoders.instEncoderScaleM2.CablePosM >= (GVL_PERSISTENT.CableLimitAscentM2_M + M2_LimitShift))
                             AND NOT PRG_04_Modes.instModes.HomingApproachEnable;

ForbidAscentM2_Raw  := PRG_03_Safety.instSafetyWinchM2.ForbidAscent
                       OR (PRG_02_Encoders.instHomingM2.Homed
                           AND NOT PRG_02_Encoders.instHomingM2.HomingSuspect
                           AND (PRG_02_Encoders.instEncoderScaleM2.CablePosM >= (GVL_PERSISTENT.HomingTargetM2_M + M2_LimitShift)))
                       OR CableLimitAscentM2Reached;

SafeStopM1_Active      := SafeStopM1_Raw      OR (instWinchSync.SyncActive AND SafeStopM2_Raw);
SafeStopM2_Active      := SafeStopM2_Raw      OR (instWinchSync.SyncActive AND SafeStopM1_Raw);
ForbidDescentM1_Active := ForbidDescentM1_Raw OR (instWinchSync.SyncActive AND ForbidDescentM2_Raw);
ForbidDescentM2_Active := ForbidDescentM2_Raw OR (instWinchSync.SyncActive AND ForbidDescentM1_Raw);
ForbidAscentM1_Active  := ForbidAscentM1_Raw  OR (instWinchSync.SyncActive AND ForbidAscentM2_Raw);
ForbidAscentM2_Active  := ForbidAscentM2_Raw  OR (instWinchSync.SyncActive AND ForbidAscentM1_Raw);

// ── 6. EXÉCUTION DU PILOTAGE DU TREUIL M1 ───────────────────────────────
instWinchM1(
    Enable                  := StubMachineEnableN1 AND NOT PRG_04_Modes.instModes.InhibitM1, // 🆕 REX 2026-07-08
    Reset                   := PRG_09_Supervision.FaultMachineReset_IHM,
    EmergencyStopOk         := PRG_00_Inputs.EmergencyStopOk,
    Mode                    := PRG_04_Modes.instModes.Mode,
    StartStop               := M1_StartStop_Active,
    SafeStop                := SafeStopM1_Active,
    ForbidDescent           := ForbidDescentM1_Active,
    ForbidAscent            := ForbidAscentM1_Active,
    Direction               := M1_Direction_Active,
    SpeedRefPct             := M1_SpeedRef_Active,
    SpeedStepTable          := GVL_PERSISTENT.WinchSpeedStepTable,
    // 🔧 REX 2026-07-15 (9) : EffectiveMaxStepDescente/Ascent (voir calcul plus haut) — Auto garde
    // WinchMaxStepDescente/5 inchangés, Manu applique en plus WinchMaxStepFwd/Rev (essais progressifs).
    MaxStepDescente         := EffectiveMaxStepDescente,
    MaxStepAscent           := EffectiveMaxStepAscent,
    HomingApproachActive    := PRG_04_Modes.instModes.HomingApproachEnable, // 🆕 REX 2026-07-08 : vitesse lente en approche
    FwdRevSpeedFeedbackOff  := PRG_00_Inputs.M1FwdRevSpeedFeedbackOff, // 🔧 REX 2026-07-07
    BrakeFeedback           := PRG_00_Inputs.M1BrakeFeedback,
    BypassContactorCheck    := GVL_Simulation.SimulationModeActive AND NOT GVL_Simulation.ContactorFeedbackM1_IsReal,
    RampAccelRate           := GVL_PERSISTENT.WinchM1RampAccelRate_Pct,
    RampDecelNormalRate     := GVL_PERSISTENT.WinchM1RampDecelNormal_Pct,
    RampDecelFastRate       := GVL_PERSISTENT.WinchM1RampDecelFast_Pct,
    Homed                   := PRG_02_Encoders.instHomingM1.Homed,
    HomingSuspect           := PRG_02_Encoders.instHomingM1.HomingSuspect, // 🆕 Câblage de l'incertitude M1
    CablePosM               := PRG_02_Encoders.instEncoderScaleM1.CablePosM,
    // 🔧 REX 2026-07-15 (6) : CableLimitAscentM1_M (limite ABSOLUE d'exploitation normale, ex-
    // HomingTargetM1_M) — la rampe/ralentissement de FB_Winch cible désormais la même limite que
    // ForbidAscentM1_Raw ci-dessus, pas le capteur physique (réservé au Homing).
    TopLimitM               := GVL_PERSISTENT.CableLimitAscentM1_M,
    BottomLimitM            := BottomLimitM1_Active,
    SlowdownDistanceM       := GVL_PERSISTENT.WinchSlowdownDistance_M,
    SlowSpeedPct            := GVL_PERSISTENT.WinchSlowSpeedPct
);

// ── 7. EXÉCUTION DU PILOTAGE DU TREUIL M2 ───────────────────────────────
instWinchM2(
    Enable                  := StubMachineEnableN1 AND NOT PRG_04_Modes.instModes.InhibitM2, // 🆕 REX 2026-07-08
    Reset                   := PRG_09_Supervision.FaultMachineReset_IHM,
    EmergencyStopOk         := PRG_00_Inputs.EmergencyStopOk,
    Mode                    := PRG_04_Modes.instModes.Mode,
    StartStop               := M2_StartStop_Active,
    SafeStop                := SafeStopM2_Active,
    ForbidDescent           := ForbidDescentM2_Active,
    ForbidAscent            := ForbidAscentM2_Active,
    Direction               := M2_Direction_Active,
    SpeedRefPct             := M2_SpeedRef_Active,
    SpeedStepTable          := M2_SpeedStepTableActive,
    // 🔧 REX 2026-07-15 (9) : idem M1 (voir §6 ci-dessus).
    MaxStepDescente         := EffectiveMaxStepDescente,
    MaxStepAscent           := EffectiveMaxStepAscent,
    HomingApproachActive    := PRG_04_Modes.instModes.HomingApproachEnable, // 🆕 REX 2026-07-08 : vitesse lente en approche
    FwdRevSpeedFeedbackOff  := PRG_00_Inputs.M2FwdRevSpeedFeedbackOff, // 🔧 REX 2026-07-07
    BrakeFeedback           := PRG_00_Inputs.M2BrakeFeedback,
    BypassContactorCheck    := GVL_Simulation.SimulationModeActive AND NOT GVL_Simulation.ContactorFeedbackM2_IsReal,
    RampAccelRate           := GVL_PERSISTENT.WinchM2RampAccelRate_Pct,
    RampDecelNormalRate     := GVL_PERSISTENT.WinchM2RampDecelNormal_Pct,
    RampDecelFastRate       := GVL_PERSISTENT.WinchM2RampDecelFast_Pct,
    Homed                   := PRG_02_Encoders.instHomingM2.Homed,
    HomingSuspect           := PRG_02_Encoders.instHomingM2.HomingSuspect, // 🆕 Câblage de l'incertitude M2
    CablePosM               := PRG_02_Encoders.instEncoderScaleM2.CablePosM,
    // 🔧 REX 2026-07-15 (6) : idem M1 (voir ci-dessus), + M2_LimitShift (décalage grappin fermé).
    TopLimitM               := GVL_PERSISTENT.CableLimitAscentM2_M + M2_LimitShift,
    BottomLimitM            := BottomLimitM2_Active,
    SlowdownDistanceM       := GVL_PERSISTENT.WinchSlowdownDistance_M,
    SlowSpeedPct            := GVL_PERSISTENT.WinchSlowSpeedPct
);

// ── 8. ALIMENTATION PRG_10_Outputs (sorties physiques) ──────────────────
// 🔴🔧 REX 2026-07-07 : PRG_10_Outputs est une tâche indépendante (MainTask, PouList),
// jamais appelée avec paramètres — ses VAR_INPUT restaient à FALSE en permanence, y compris
// sur machine réelle (aucun relais/contacteur/frein ne s'activait jamais). Alimentation directe
// ici, AVANT PRG_10_Outputs dans l'ordre de tâche (position 6 < 10, même cycle API).
PRG_10_Outputs.M1RelayFwd        := instWinchM1.RelayFwd;
PRG_10_Outputs.M1RelayRev        := instWinchM1.RelayRev;
PRG_10_Outputs.M1SpeedContactor1 := instWinchM1.Contactor1;
PRG_10_Outputs.M1SpeedContactor2 := instWinchM1.Contactor2;
PRG_10_Outputs.M1SpeedContactor3 := instWinchM1.Contactor3;
PRG_10_Outputs.M1SpeedContactor4 := instWinchM1.Contactor4;
PRG_10_Outputs.M1BrakeCmd        := instWinchM1.BrakeCmd;

PRG_10_Outputs.M2RelayFwd        := instWinchM2.RelayFwd;
PRG_10_Outputs.M2RelayRev        := instWinchM2.RelayRev;
PRG_10_Outputs.M2SpeedContactor1 := instWinchM2.Contactor1;
PRG_10_Outputs.M2SpeedContactor2 := instWinchM2.Contactor2;
PRG_10_Outputs.M2SpeedContactor3 := instWinchM2.Contactor3;
PRG_10_Outputs.M2SpeedContactor4 := instWinchM2.Contactor4;
PRG_10_Outputs.M2BrakeCmd        := instWinchM2.BrakeCmd;

(* ---- PRG_07_ChariotControl.st ---- *)
(* ═══════════════════════════════════════════════════════════════
   ↔️ PRG_07_ChariotControl — Pilotage de la Translation Chariot M3
   ───────────────────────────────────────────────────────────────
   ⚙️ Exécuté par la tâche PLC en position 7.
   ✅ Arbitre entre les commandes Manuelles (Joystick) et Automatiques (PRG_05_Cycle).
   ═══════════════════════════════════════════════════════════════ *)

PROGRAM PRG_07_ChariotControl
VAR
    instChariotM3           : FB_Chariot;

    // Commandes arbitrées après sélection Manuel/Auto
    M3_StartStop_Active     : BOOL;
    M3_Direction_Active     : INT;
    M3_SpeedRef_Active      : REAL;
    M3_PositionSensorTarget : BOOL;

    // Target active (HMI en manuel, instCycle en auto)
    SelectedTargetNum       : INT;
END_VAR

// === IMPLEMENTATION (corps du PROGRAM PRG_07_ChariotControl) ===

// ── 1. ARBITRAGE DU SÉLECTEUR DE CIBLE ET DE LA DIRECTION ──────────────────
IF PRG_04_Modes.instModes.Mode = E_Mode.SEMI_AUTO THEN
    // Mode Auto/Semi-Auto : Consigne issue du séquenceur de cycle
    SelectedTargetNum    := PRG_05_Cycle.instCycle.CmdChariotM3_Target;
    M3_StartStop_Active  := PRG_05_Cycle.instCycle.CmdChariotM3_Start;
    M3_SpeedRef_Active   := 40.0; // Vitesse de translation automatique nominale (40%)

    // Détermination automatique du sens de marche selon la cible :
    // - Trémie (cible 4) = Marche Avant (Direction := 1)
    // - Fosses (cible 1 et 2) = Marche Arrière (Direction := -1)
    IF SelectedTargetNum = 4 THEN
        M3_Direction_Active := 1;
    ELSE
        M3_Direction_Active := -1;
    END_IF;
ELSE
    // Mode Manuel/Maintenance : Consignes issues du Joystick et sélecteur HMI
    SelectedTargetNum    := StubChariotPositionSelect_IHM;
    M3_StartStop_Active  := PRG_01_Diagnostics.FB_Joystick_0.AxisCmdX.StartStop;
    M3_Direction_Active  := PRG_01_Diagnostics.FB_Joystick_0.AxisCmdX.Direction;
    M3_SpeedRef_Active   := PRG_01_Diagnostics.FB_Joystick_0.AxisCmdX.SpeedRef;
END_IF;

// Câblage du capteur de butée de la cible sélectionnée
CASE SelectedTargetNum OF
    1: M3_PositionSensorTarget := PRG_00_Inputs.ChariotPosFosse1;
    2: M3_PositionSensorTarget := PRG_00_Inputs.ChariotPosFosse2;
    3: M3_PositionSensorTarget := PRG_00_Inputs.ChariotPosMaintenance;
    4: M3_PositionSensorTarget := PRG_00_Inputs.ChariotPosTremie;
ELSE
    M3_PositionSensorTarget := FALSE;   // Aucun capteur visé
END_CASE;

// ── 2. EXÉCUTION DU PILOTAGE DU CHARIOT M3 ──────────────────────────────
instChariotM3(
    Enable                  := PRG_06_WinchControl.StubMachineEnableN1,
    Reset                   := PRG_09_Supervision.FaultMachineReset_IHM,
    EmergencyStopOk         := PRG_00_Inputs.EmergencyStopOk,
    Mode                    := PRG_04_Modes.instModes.Mode,
    StartStop               := M3_StartStop_Active,
    SafeStop                := PRG_03_Safety.instSafetyChariotM3.SafeStop,
    Direction               := M3_Direction_Active,
    SpeedRefPct             := M3_SpeedRef_Active,
    PositionSensorTarget    := M3_PositionSensorTarget,
    LimitSwitchFwd          := PRG_00_Inputs.ChariotPosTremie,
    LimitSwitchRev          := PRG_00_Inputs.ChariotPosFosse1,
    DriveStatusWord         := PRG_00_Inputs.M3_StatusWord_Filtered,
    DriveActualFreqHz       := UINT_TO_REAL(PRG_00_Inputs.M3_ActualFrequencyHz_Filtered) / 100.0,
    BrakeFeedback           := SEL(GVL_IHM.ChariotM3.BypassContactorFeedback, PRG_00_Inputs.M3BrakeFeedback, instChariotM3.BrakeCmd),
    BypassContactorCheck    := GVL_Simulation.SimulationModeActive AND NOT GVL_Simulation.ContactorFeedbackM3_IsReal
);

// 🔴 Recopie commande de frein chariot
PRG_10_Outputs.ChariotBrakeCmd := instChariotM3.BrakeCmd;

(* ---- PRG_08_AuxiliaryControl.st ---- *)
(* ═══════════════════════════════════════════════════════════════
   ⚡ PRG_08_AuxiliaryControl — Gestion des Auxiliaires (Hydraulique, Crible...)
   ───────────────────────────────────────────────────────────────
   ⚙️ Exécuté par la tâche PLC en position 8.
   ✅ Regroupe toutes les commandes et logiques hors-axes.
   ═══════════════════════════════════════════════════════════════ *)

PROGRAM PRG_08_AuxiliaryControl
VAR_INPUT
    // 🌡️ Groupe Hydraulique
    HydraulicPumpRunCmd   : BOOL;   // Commande démarrage centrale hydraulique
    HydraulicFaultOk      : BOOL;   // Retour défaut groupe hydraulique (NC)

    // 🌾 Crible (Sifter / Sieve)
    SifterRunCmd          : BOOL;   // Commande marche crible
    SifterFaultOk         : BOOL;   // Retour défaut électrique crible (NC)

    // 🔗 Divers
    GridOpenCmd           : BOOL;   // Commande ouverture grille
    HelmetCloseCmd        : BOOL;   // Commande fermeture casque
END_VAR

// === IMPLEMENTATION (corps du PROGRAM PRG_08_AuxiliaryControl) ===

// --- STUBS LOGIQUES TEMPORAIRES (comportement passif / neutre) ---
// HydraulicPumpRunCmd := FALSE; // Commenté pour permettre le pilotage externe (ex: PRG_10_Outputs)
// SifterRunCmd        := FALSE;
// GridOpenCmd         := FALSE;
// HelmetCloseCmd      := FALSE;

HydraulicFaultOk    := TRUE; // Par défaut sain (NC)
SifterFaultOk       := TRUE; // Par défaut sain (NC)
